(* IEC 61131-3 sources: JingjiangArm/moonboxpro_arm_8.4/Application/Application/任务列表/TensionTask/电机运动/MotionCtl_GantryTrap (part 2) *)

		//如果版辊周长变了/料膜厚度变了2023.12.27.171307
		IF (pstStGrpParam_Save^.rFilmThick_Confirm<>pstStGrpParam_Save^.rFilmThickNess_Using AND
			pstStGrpParam_Save^.rFilmThick_Confirm<>0 AND pstStGrpParam_Save^.rFilmThickNess_Using<>0) OR
			pstStUnitParam_Save^.rGirth_Confirmed_press_dn_NetRoller<>pstStUnitParam_Save^.rGirth_NetRoller OR
			pstStUnitParam_Save^.rGirth_Confirmed_press_dn_PrnRoller<>pstStUnitParam_Save^.rGirth_PrnRoller OR
			rGirth_PrnRoller_Mem <> pstStGrpParam_Save^.rGirth_PrnRoller THEN
			//处理一下位置更新2023.12.27.171801
			lrTemp:= g_rPos_press_dn_NetRoller_Pressure_MM*GC_LRMOTORPPR_TRAP*
						UINT_TO_REAL(pstStUnitParam_Save^.uiNum_NetRoller_Pressure)/
						pstStUnitParam_Save^.rScrewPitch_NetRoller_Pressure/
						UINT_TO_REAL(pstStUnitParam_Save^.uiDen_NetRoller_Pressure);

			IF i_pastStTrapAxisParam_Gantray^[2,iN].xRev_Motor_M THEN

				i_pastStTrapAxisParam_Gantray^[2,iN].lrposConfirm_Dn_Press_M:= i_pastStTrapAxisParam_Gantray^[2,iN].lrposConfirm_Dn_Press_M_Confirm-
						((
						(pstStGrpParam_Save^.rFilmThick_Manu-pstStGrpParam_Save^.rFilmThick_Confirm))*
						UINT_TO_LREAL(pstStUnitParam_Save^.uiNum_NetRoller_Pressure)*GC_LRMOTORPPR_TRAP/
						UINT_TO_LREAL(pstStUnitParam_Save^.uiDen_NetRoller_Pressure)/pstStUnitParam_Save^.rScrewPitch_NetRoller_Pressure);

				i_pastStTrapAxisParam_Gantray^[2,iN].lrposConfirm_Up_Press_M:= i_pastStTrapAxisParam_Gantray^[2,iN].lrposConfirm_Dn_Press_M-lrTemp;
			ELSE

					i_pastStTrapAxisParam_Gantray^[2,iN].lrposConfirm_Dn_Press_M:= i_pastStTrapAxisParam_Gantray^[2,iN].lrposConfirm_Dn_Press_M_Confirm+
						((
						(pstStGrpParam_Save^.rFilmThick_Manu-pstStGrpParam_Save^.rFilmThick_Confirm))*
						UINT_TO_LREAL(pstStUnitParam_Save^.uiNum_NetRoller_Pressure)*GC_LRMOTORPPR_TRAP/
						UINT_TO_LREAL(pstStUnitParam_Save^.uiDen_NetRoller_Pressure)/pstStUnitParam_Save^.rScrewPitch_NetRoller_Pressure);

				i_pastStTrapAxisParam_Gantray^[2,iN].lrposConfirm_Up_Press_M:= i_pastStTrapAxisParam_Gantray^[2,iN].lrposConfirm_Dn_Press_M+lrTemp;
			END_IF
			IF i_pastStTrapAxisParam_Gantray^[2,iN].xRev_Motor_G THEN

				i_pastStTrapAxisParam_Gantray^[2,iN].lrposConfirm_Dn_Press_G:= i_pastStTrapAxisParam_Gantray^[2,iN].lrposConfirm_Dn_Press_G_Confirm-
						(((*(i_pastStTrapAxisParam_Gantray^[2,iN].rweigth_Zero-
						i_pastStTrapAxisParam_Gantray^[2,iN].rweigth_Zero_Confirm)+*)
						(pstStGrpParam_Save^.rFilmThickNess_Using-pstStGrpParam_Save^.rFilmThick_Confirm))*
						UINT_TO_LREAL(pstStUnitParam_Save^.uiNum_NetRoller_Pressure)*GC_LRMOTORPPR_TRAP/
						UINT_TO_LREAL(pstStUnitParam_Save^.uiDen_NetRoller_Pressure)/pstStUnitParam_Save^.rScrewPitch_NetRoller_Pressure);
				i_pastStTrapAxisParam_Gantray^[2,iN].lrposConfirm_Up_Press_G:= i_pastStTrapAxisParam_Gantray^[2,iN].lrposConfirm_Dn_Press_G-lrTemp;
			ELSE

					i_pastStTrapAxisParam_Gantray^[2,iN].lrposConfirm_Dn_Press_G:= i_pastStTrapAxisParam_Gantray^[2,iN].lrposConfirm_Dn_Press_G_Confirm+
							(((i_pastStTrapAxisParam_Gantray^[2,iN].rweigth_Zero-
							i_pastStTrapAxisParam_Gantray^[2,iN].rweigth_Zero_Confirm)+
							(pstStGrpParam_Save^.rFilmThick_Manu-pstStGrpParam_Save^.rFilmThick_Confirm))*
							UINT_TO_LREAL(pstStUnitParam_Save^.uiNum_NetRoller_Pressure)*GC_LRMOTORPPR_TRAP/
							UINT_TO_LREAL(pstStUnitParam_Save^.uiDen_NetRoller_Pressure)/pstStUnitParam_Save^.rScrewPitch_NetRoller_Pressure);

				i_pastStTrapAxisParam_Gantray^[2,iN].lrposConfirm_Up_Press_G:= i_pastStTrapAxisParam_Gantray^[2,iN].lrposConfirm_Dn_Press_G+lrTemp;
			END_IF
			i_pastStTrapAxisParam_Gantray^[2,iN].lrposConfirm_Load_Unload_Press_M:= //换版位的物理位置是不变的2023.12.13.081145
				i_pastStTrapAxisParam_Gantray^[2,iN].lrposConfirm_Load_Unload_Press_M_Confirm;
			i_pastStTrapAxisParam_Gantray^[2,iN].lrposConfirm_Load_Unload_Press_G:=
				i_pastStTrapAxisParam_Gantray^[2,iN].lrposConfirm_Load_Unload_Press_G_Confirm;
		ELSE
			//bai.zy | 2024.03.21.130939 | 增加印刷位
			i_pastStTrapAxisParam_Gantray^[2,iN].lrposConfirm_Dn_Press_M:=
				i_pastStTrapAxisParam_Gantray^[2,iN].lrposConfirm_Dn_Press_M_Confirm;
			i_pastStTrapAxisParam_Gantray^[2,iN].lrposConfirm_Dn_Press_G:=
				i_pastStTrapAxisParam_Gantray^[2,iN].lrposConfirm_Dn_Press_G_Confirm;
			i_pastStTrapAxisParam_Gantray^[2,iN].lrposConfirm_Up_Press_M:=
				i_pastStTrapAxisParam_Gantray^[2,iN].lrposConfirm_Up_Press_M_Confirm;
			i_pastStTrapAxisParam_Gantray^[2,iN].lrposConfirm_Up_Press_G:=
				i_pastStTrapAxisParam_Gantray^[2,iN].lrposConfirm_Up_Press_G_Confirm;
			i_pastStTrapAxisParam_Gantray^[2,iN].lrposConfirm_Load_Unload_Press_M:= //换版位的物理位置是不变的2023.12.13.081145
				i_pastStTrapAxisParam_Gantray^[2,iN].lrposConfirm_Load_Unload_Press_M_Confirm;
			i_pastStTrapAxisParam_Gantray^[2,iN].lrposConfirm_Load_Unload_Press_G:=
				i_pastStTrapAxisParam_Gantray^[2,iN].lrposConfirm_Load_Unload_Press_G_Confirm;

		END_IF
	//2026.02.07.160105 计算网辊步进量

		afbKS_FB_GantryTrap_Calc_TargetPos_Net[iN](
			i_xEn:= TRUE,
			i_uiNum:= pstStUnitParam_Save^.uiNum_NetRoller_Pressure,
			i_uiDen:= pstStUnitParam_Save^.uiDen_NetRoller_Pressure,
			i_rScrewPitch:= pstStUnitParam_Save^.rScrewPitch_NetRoller_Pressure,
			i_rUp_Dn_Length:= g_rPos_press_dn_NetRoller_Pressure_MM,//1.35, //3mm
			i_rGirth_Roller:= pstStUnitParam_Save^.rGirth_NetRoller,
			i_xStopOrEstop_Valid:= xNeedMoveUp_Stop_Net,
			i_prGirth_Confirm:= ADR(pstStUnitParam_Save^.rGirth_Confirmed_press_dn_NetRoller),
			i_xFlag_Print:= pstStGrpParam_UnSave^.xFlag_Print,
			i_xStep_Fast:= pstStUnitParam_Save^.wFlag_PressFun.2,//^.xStep_Fast,
			i_rStep_Fast:= pstStGrpParam_Save^.rStep_Fast,
			i_rStep_Little:= pstStGrpParam_Save^.rStep_Little,
			i_rVel_Fast:= pstStGrpParam_Save^.rVel_Press_Net,//
			i_rVel_Little:= 0.1,
			i_plrTargetPos_All:= ADR(alrTargetPos_Net[iN]),
			i_plrTargetPos_M:= ADR(alrTargetPos_Net_M[iN]),
			i_plrTargetPos_G:= ADR(alrTargetPos_Net_G[iN]),
			i_pstStTrapAxisParam_Gantray:= ADR(i_pastStTrapAxisParam_Gantray^[2,iN]),
			i_xFlag_Estop:= i_xFlag_Estop,
			//i_rStep_HMI:= pstStUnitParam^.rStep_Pressure_Prn_Net,//2023.12.22.220303
			//i_rDistanceForAvoidPrnGear := 0,
			i_pxFinishConfirm_Adjust_PressDn := ADR(axFinishConfirm_Adjust_PressDn[iN]),//: POINTER TO BOOL;
			i_rStep_HMI_Use:=pstStUnitParam_Save^.rStep_Pressure_Prn_Net,
			i_rProportion:=1.0,
			i_xMove_to_Up_Estop := pstStGrpParam_Save^.wCtl_Pressure_Up_Dn.1,
			i_ReqResetEstop := i_ReqResetEstop,
			i_rMaxErr := rMaxErr,
			o_xEn=> ,
			o_rVel=> o_arVel_Net[iN],
			o_lrTargetPos_All=> o_alrTargetPos_Net[iN],
			o_lrTargetPos_M=> o_alrTargetPos_Net_M[iN],
			o_lrTargetPos_G=> o_alrTargetPos_Net_G[iN],
			o_lrTemp_Len_Up_Pos=>alrTemp_Len_Up_Pos_Net[iN],
			o_lrTemp_Len_Load_Unload_Pos=>alrTemp_Len_Load_Unload_Pos_Net[iN]);

		pstStUnitParam_Save^.rPos_load_unload_NetRoller_Pressure_M:=
			i_pastStTrapAxisParam_Gantray^[2,iN].lrposConfirm_Load_Unload_Press_M_Confirm;
		pstStUnitParam_Save^.rPos_load_unload_NetRoller_Pressure_G:=
			i_pastStTrapAxisParam_Gantray^[2,iN].lrposConfirm_Load_Unload_Press_G_Confirm;
		pstStUnitParam_Save^.rPos_press_up_NetRoller_Pressure_M:=
			i_pastStTrapAxisParam_Gantray^[2,iN].lrposConfirm_Up_Press_M_Confirm;
		pstStUnitParam_Save^.rPos_press_up_NetRoller_Pressure_G:=
			i_pastStTrapAxisParam_Gantray^[2,iN].lrposConfirm_Up_Press_G_Confirm;
		pstStUnitParam_Save^.rPos_press_dn_NetRoller_Pressure_M:=
			i_pastStTrapAxisParam_Gantray^[2,iN].lrposConfirm_Dn_Press_M_Confirm;
		pstStUnitParam_Save^.rPos_press_dn_NetRoller_Pressure_G:=
			i_pastStTrapAxisParam_Gantray^[2,iN].lrposConfirm_Dn_Press_G_Confirm;
		pstStUnitParam_UnSave^.rPos_NetRoller_Pressure_M:= LREAL_TO_REAL(i_pastStTrapAxisParam_Gantray^[2,iN].lrCurPos_mm_M);
		pstStUnitParam_UnSave^.rPos_NetRoller_Pressure_G:= LREAL_TO_REAL(i_pastStTrapAxisParam_Gantray^[2,iN].lrCurPos_mm_G);

		//bai.zy | 2024.01.15.105513 | 合压位换版位标定完成标志
		pstStUnitParam_Save^.xConfirmDnPosDne_NetRoller_Pressure_M := i_pastStTrapAxisParam_Gantray^[2,iN].xConfirmDnPosDne_Pressure_M;
		pstStUnitParam_Save^.xConfirmDnPosDne_NetRoller_Pressure_G := i_pastStTrapAxisParam_Gantray^[2,iN].xConfirmDnPosDne_Pressure_G;
		pstStUnitParam_Save^.xConfirmload_unloadPosDne_NetRoller_Pressure_M := i_pastStTrapAxisParam_Gantray^[2,iN].xConfirmload_unloadPosDne_Pressure_M;
		pstStUnitParam_Save^.xConfirmload_unloadPosDne_NetRoller_Pressure_G := i_pastStTrapAxisParam_Gantray^[2,iN].xConfirmload_unloadPosDne_Pressure_G;

		//2024.10.21.121704
		IF pstStUnitParam_UnSave^.xConfirmParallelPos_Net THEN//平行确认按钮
			pstStUnitParam_Save^.axPressLimit_Min[2] := TRUE;
			pstStUnitParam_Save^.lrEncPosParallel_Net_M:=i_pastStTrapAxisParam_Gantray^[2,iN].lrEncPosParallel_M;//平行编码器值
			pstStUnitParam_Save^.lrEncPosParallel_Net_G:=i_pastStTrapAxisParam_Gantray^[2,iN].lrEncPosParallel_G;
			pstStUnitParam_UnSave^.xConfirmParallelPos_Net := FALSE;
		END_IF
		pstStUnitParam_UnSave^.rParallelError_Net_MM := i_pastStTrapAxisParam_Gantray^[2,iN].lrParallelError_MM;
		pstStUnitParam_Save^.lrPrintPosOffsetDn_Net_M:=i_pastStTrapAxisParam_Gantray^[2,iN].lrPrintPosOffsetDn_M;//合压偏移量
		pstStUnitParam_Save^.lrPrintPosOffsetDn_Net_G:=i_pastStTrapAxisParam_Gantray^[2,iN].lrPrintPosOffsetDn_G;

		IF pstStUnitParam_UnSave^.axCalidPressLimit_Max[2] THEN
			pstStUnitParam_UnSave^.axCalidPressLimit_Max[2] := FALSE;
			pstStUnitParam_Save^.axPressLimit_Max[2] := TRUE;
			pstStUnitParam_Save^.lrEncPosLimit_Net_M_Max := i_pastStTrapAxisParam_Gantray^[2,iN].lrEncPosLimit_M_Max ;
			pstStUnitParam_Save^.lrEncPosLimit_Net_G_Max := i_pastStTrapAxisParam_Gantray^[2,iN].lrEncPosLimit_G_Max ;
		END_IF

	END_FOR

	//版周长

	rGirth_PrnRoller_Mem := pstStGrpParam_Save^.rGirth_PrnRoller;		//	秦华不需要了

	FOR iN:=1 TO i_iGrpUnitNum_Pu BY 1 DO
		IF axFlag_Mode_Calid[iN] THEN
			g_xModeCalibSwitch_Flag := TRUE;
			IF NOT i_xDebugMode THEN
				g_xModeCalibSwitch_Flag := FALSE;
			END_IF
			EXIT;
		ELSE
			g_xModeCalibSwitch_Flag := FALSE;
		END_IF
	END_FOR

	IF i_xDebugMode THEN
		FOR iN := 1 TO i_iGrpUnitNum_Pu BY 1 DO
			pstStUnitParam_Save:= ADR(i_pstStSysParam^.astStUnitParam_Save[iN]);
			pstStUnitParam_UnSave:= ADR(i_pstStSysParam^.astStUnitParam_UnSave[iN]);
			axTRIG_ResetFlag_FinishCalid[iN](CLK:=g_axResetFlag_FinishCalid[iN]);
			IF axTRIG_ResetFlag_FinishCalid[iN].Q THEN
				g_axResetFlag_FinishCalid[iN] := FALSE;

				pstStUnitParam_Save^.xConfirmDnPosDne_PrnRoller_Pressure_M:=FALSE;
				pstStUnitParam_Save^.xConfirmDnPosDne_PrnRoller_Pressure_G:=FALSE;
				pstStUnitParam_Save^.xConfirmDnPosDne_NetRoller_Pressure_M:=FALSE;
				pstStUnitParam_Save^.xConfirmDnPosDne_NetRoller_Pressure_G:=FALSE;
				pstStUnitParam_Save^.xConfirmload_unloadPosDne_PrnRoller_Pressure_M:=FALSE;
				pstStUnitParam_Save^.xConfirmload_unloadPosDne_PrnRoller_Pressure_G:=FALSE;
				pstStUnitParam_Save^.xConfirmload_unloadPosDne_NetRoller_Pressure_M:=FALSE;
				pstStUnitParam_Save^.xConfirmload_unloadPosDne_NetRoller_Pressure_G:=FALSE;

				pstStUnitParam_Save^.xConfirmDnPosDne_StrRoller_Pressure_M:=FALSE;
				pstStUnitParam_Save^.xConfirmDnPosDne_StrRoller_Pressure_G:=FALSE;
				//印版
				pstStUnitParam_Save^.rPos_load_unload_PrnRoller_Pressure_M := 0;//换版位
				pstStUnitParam_Save^.rPos_load_unload_PrnRoller_Pressure_G := 0;
				pstStUnitParam_Save^.rPos_press_up_PrnRoller_Pressure_M := 0;//离压位
				pstStUnitParam_Save^.rPos_press_up_PrnRoller_Pressure_G := 0;
				pstStUnitParam_Save^.rPos_press_dn_PrnRoller_Pressure_M := 0;//合压位
				pstStUnitParam_Save^.rPos_press_dn_PrnRoller_Pressure_G := 0;
				pstStUnitParam_Save^.liABSPos_Prn_M := 0;
				pstStUnitParam_Save^.liABSPos_Prn_G := 0;
				//网辊
				pstStUnitParam_Save^.rPos_load_unload_NetRoller_Pressure_M := 0;//换版位
				pstStUnitParam_Save^.rPos_load_unload_NetRoller_Pressure_G := 0;
				pstStUnitParam_Save^.rPos_press_up_NetRoller_Pressure_M := 0;//离压位
				pstStUnitParam_Save^.rPos_press_up_NetRoller_Pressure_G := 0;
				pstStUnitParam_Save^.rPos_press_dn_NetRoller_Pressure_M := 0;//合压位
				pstStUnitParam_Save^.rPos_press_dn_NetRoller_Pressure_G := 0;
				pstStUnitParam_Save^.liABSPos_Net_M := 0;
				pstStUnitParam_Save^.liABSPos_Net_G := 0;
				//张带
				pstStUnitParam_Save^.rPos_load_unload_StrRoller_Pressure_M := 0;//换版位
				pstStUnitParam_Save^.rPos_load_unload_StrRoller_Pressure_G := 0;
				pstStUnitParam_Save^.rPos_press_up_StrRoller_Pressure_M := 0;//离压位
				pstStUnitParam_Save^.rPos_press_up_StrRoller_Pressure_G := 0;
				pstStUnitParam_Save^.rPos_press_dn_StrRoller_Pressure_M := 0;//合压位
				pstStUnitParam_Save^.rPos_press_dn_StrRoller_Pressure_G := 0;
				pstStUnitParam_Save^.liABSPos_Str_M := 0;
				pstStUnitParam_Save^.liABSPos_Str_G := 0;

				FOR iM := 1 TO gc_iMax_PressureRoller_Unit BY 1 DO
					aitargetStation[2*iM-1] := (i_pastStTrapAxisParam_Gantray^[iM,iN].iStationId_M);
					aitargetStation[2*iM] := (i_pastStTrapAxisParam_Gantray^[iM,iN].iStationId_G);
					aliABSEncPos[2*iM-1] := 0;
					aliABSEncPos[2*iM] := 0;
				END_FOR
				//iRtn := GT_RN_SetTrapCoordinate(targetNum:= INT_TO_BYTE(gc_iMax_PressureRoller_Unit*2), targetStation:= ADR(abytargetStation), targetAxis:= ADR(aliABSEncPos));

				axAxisRev[1]:= i_pastStTrapAxisParam_Gantray^[1,iN].xRev_Motor_M;
				axAxisRev[2]:= i_pastStTrapAxisParam_Gantray^[1,iN].xRev_Motor_G;
				axAxisRev[3]:= i_pastStTrapAxisParam_Gantray^[2,iN].xRev_Motor_M;
				axAxisRev[4]:= i_pastStTrapAxisParam_Gantray^[2,iN].xRev_Motor_G;
				axAxisRev[5]:= i_pastStTrapAxisParam_Gantray^[3,iN].xRev_Motor_M;
				axAxisRev[6]:= i_pastStTrapAxisParam_Gantray^[3,iN].xRev_Motor_G;

				iRtn := KS_SetTrapCoordinate(
						i_xEn:= TRUE,
						i_iTarget_Num:= INT_TO_BYTE(gc_iMax_PressureRoller_Unit*2),
						i_paiTargetStationList:= ADR(aitargetStation),
						i_paliABSEncPos:= ADR(aliABSEncPos),
						i_paxAxisRev:= ADR(axAxisRev),
						i_pastStAxisIdListInf:= i_pastStAxisIdListInf,
						i_pastStGetMotionSts:= i_pastStGetMotionSts,
						i_pstStSysStationInf := i_pstStSysStationInf,
						i_pstStSysGantryAxisInf := i_pstStSysGantryAxisInf,
						ADR(g_alrCurrentAbsPos_Debug));

			END_IF
		END_FOR
	END_IF

(*
	FOR iN := 1 TO i_iGrpUnitNum_Pu BY 1 DO
		pstStUnitParam_Save:= ADR(i_pstStSysParam^.astStUnitParam_Save[iN]);
		pstStUnitParam_UnSave:= ADR(i_pstStSysParam^.astStUnitParam_UnSave[iN]);
		//印刷过程中矫正合压位是否要重新清零清规划？？？？
		//矫正后更新当前参数值
		//2025.08.28.152652 | 矫正增加对于压力电机的位置判断，之前做过判断，但是不再范围内的位置还是被矫正了，这里再次判断一下
		IF axFinishConfirm_Adjust_PressDn[iN] AND
			pstStUnitParam_Save^.xLinkage AND
			(i_pastStTrapAxisParam_Gantray^[1,iN].byCurPos_M = 1 OR
			i_pastStTrapAxisParam_Gantray^[1,iN].byCurPos_M = 2 OR
			i_pastStTrapAxisParam_Gantray^[1,iN].byCurPos_M = 3 ) AND
			(i_pastStTrapAxisParam_Gantray^[1,iN].byCurPos_G = 1 OR
			i_pastStTrapAxisParam_Gantray^[1,iN].byCurPos_G = 2 OR
			i_pastStTrapAxisParam_Gantray^[1,iN].byCurPos_G = 3 ) AND
			(i_pastStTrapAxisParam_Gantray^[2,iN].byCurPos_M = 1 OR
			i_pastStTrapAxisParam_Gantray^[2,iN].byCurPos_M = 2 OR
			i_pastStTrapAxisParam_Gantray^[2,iN].byCurPos_M = 3 ) AND
			(i_pastStTrapAxisParam_Gantray^[2,iN].byCurPos_G = 1 OR
			i_pastStTrapAxisParam_Gantray^[2,iN].byCurPos_G = 2 OR
			i_pastStTrapAxisParam_Gantray^[2,iN].byCurPos_G = 3 ) THEN

			axFinishConfirm_Adjust_PressDn[iN] := FALSE;

			alrTemp_Len_Up_Pos_Prn[iN] := g_rPos_press_dn_PrnRoller_Pressure_MM(*i_pstStSysParam^.rPos_press_dn_PrnRoller_Pressure_MM*)*
										pstStUnitParam_Save^.uiNum_PrnRoller_Pressure*GC_LRMOTORPPR_TRAP/
										pstStUnitParam_Save^.uiDen_PrnRoller_Pressure/pstStUnitParam_Save^.rScrewPitch_PrnRoller_Pressure;
			alrTemp_Len_Load_Unload_Pos_Prn[iN] :=g_rPos_press_dn_PrnRoller_Pressure_MM(*i_pstStSysParam^.rPos_load_unload_PrnRoller_Pressure_MM*)*
										pstStUnitParam_Save^.uiNum_PrnRoller_Pressure*GC_LRMOTORPPR_TRAP/
										pstStUnitParam_Save^.uiDen_PrnRoller_Pressure/pstStUnitParam_Save^.rScrewPitch_PrnRoller_Pressure;
			//印版
			iRtn := GTN_RN_GetAxisAbsPosEx(cardNum:= 1, axis:= 1, pPos:= ADR(g_liAbsPos_M), stationId:= i_pastStTrapAxisParam_Gantray^[1,iN].iStationId_M);
			iRtn := GTN_RN_GetAxisAbsPosEx(cardNum:= 1, axis:= 1, pPos:= ADR(g_liAbsPos_G), stationId:= i_pastStTrapAxisParam_Gantray^[1,iN].iStationId_G);
			pstStUnitParam_Save^.rPos_press_dn_PrnRoller_Pressure_M:= 1;//LINT_TO_LREAL(g_liAbsPos_M);
			pstStUnitParam_Save^.rPos_press_dn_PrnRoller_Pressure_G:= 1;//LINT_TO_LREAL(g_liAbsPos_G);
			pstStUnitParam_Save^.rPos_press_up_PrnRoller_Pressure_M:= pstStUnitParam_Save^.rPos_press_dn_PrnRoller_Pressure_M + alrTemp_Len_Up_Pos_Prn[iN];//1;//LINT_TO_LREAL(g_liAbsPos_M);
			pstStUnitParam_Save^.rPos_press_up_PrnRoller_Pressure_G:= pstStUnitParam_Save^.rPos_press_dn_PrnRoller_Pressure_G + alrTemp_Len_Up_Pos_Prn[iN];//1;//LINT_TO_LREAL(g_liAbsPos_G);
			pstStUnitParam_Save^.rPos_load_unload_PrnRoller_Pressure_M:= pstStUnitParam_Save^.rPos_press_dn_PrnRoller_Pressure_M + alrTemp_Len_Load_Unload_Pos_Prn[iN];//1;//LINT_TO_LREAL(g_liAbsPos_M);
			pstStUnitParam_Save^.rPos_load_unload_PrnRoller_Pressure_G:= pstStUnitParam_Save^.rPos_press_dn_PrnRoller_Pressure_G + alrTemp_Len_Load_Unload_Pos_Prn[iN];//1;//LINT_TO_LREAL(g_liAbsPos_G);
			iRtn := GT_RN_SetTrapCoordinate(targetNum:=1 , targetStation:=ADR(i_pastStTrapAxisParam_Gantray^[1,iN].iStationId_M),targetAxis:= ADR(g_liAbsPos_M));
			iRtn := GT_RN_SetTrapCoordinate(targetNum:=1 , targetStation:=ADR(i_pastStTrapAxisParam_Gantray^[1,iN].iStationId_G),targetAxis:= ADR(g_liAbsPos_G));
			pstStUnitParam_Save^.liABSPos_Prn_M := g_liAbsPos_M;
			pstStUnitParam_Save^.liABSPos_Prn_G := g_liAbsPos_G;
			//网辊
			iRtn := GTN_RN_GetAxisAbsPosEx(cardNum:= 1, axis:= 1, pPos:= ADR(g_liAbsPos_M), stationId:= i_pastStTrapAxisParam_Gantray^[2,iN].iStationId_M);
			iRtn := GTN_RN_GetAxisAbsPosEx(cardNum:= 1, axis:= 1, pPos:= ADR(g_liAbsPos_G), stationId:= i_pastStTrapAxisParam_Gantray^[2,iN].iStationId_G);
			pstStUnitParam_Save^.rPos_press_dn_NetRoller_Pressure_M:= 1;//LINT_TO_LREAL(g_liAbsPos_M);
			pstStUnitParam_Save^.rPos_press_dn_NetRoller_Pressure_G:= 1;//LINT_TO_LREAL(g_liAbsPos_G);
			pstStUnitParam_Save^.rPos_press_up_NetRoller_Pressure_M:= pstStUnitParam_Save^.rPos_press_dn_NetRoller_Pressure_M + alrTemp_Len_Up_Pos_Net[iN];//1;//LINT_TO_LREAL(g_liAbsPos_M);
			pstStUnitParam_Save^.rPos_press_up_NetRoller_Pressure_G:= pstStUnitParam_Save^.rPos_press_dn_NetRoller_Pressure_G + alrTemp_Len_Up_Pos_Net[iN];//1;//LINT_TO_LREAL(g_liAbsPos_G);
			pstStUnitParam_Save^.rPos_load_unload_NetRoller_Pressure_M:= pstStUnitParam_Save^.rPos_press_dn_NetRoller_Pressure_M + alrTemp_Len_Load_Unload_Pos_Net[iN];//1;//LINT_TO_LREAL(g_liAbsPos_M);
			pstStUnitParam_Save^.rPos_load_unload_NetRoller_Pressure_G:= pstStUnitParam_Save^.rPos_press_dn_NetRoller_Pressure_G + alrTemp_Len_Load_Unload_Pos_Net[iN];//1;//LINT_TO_LREAL(g_liAbsPos_G);
			iRtn := GT_RN_SetTrapCoordinate(targetNum:=1 , targetStation:=ADR(i_pastStTrapAxisParam_Gantray^[2,iN].iStationId_M),targetAxis:= ADR(g_liAbsPos_M));
			iRtn := GT_RN_SetTrapCoordinate(targetNum:=1 , targetStation:=ADR(i_pastStTrapAxisParam_Gantray^[2,iN].iStationId_G),targetAxis:= ADR(g_liAbsPos_G));
			pstStUnitParam_Save^.liABSPos_Net_M := g_liAbsPos_M;
			pstStUnitParam_Save^.liABSPos_Net_G := g_liAbsPos_G;

		END_IF
	END_FOR
*)
IF xtest4 THEN
	xtest4:=FALSE;
	iRtn := GTN_RN_ReadAbsEncPos(cardIndex:= 1, stationPhyId:=  113, encoder:= 1, pPos:= ADR(lrAbsPos1));
	iRtn := GTN_RN_ReadAbsEncPos(cardIndex:= 1, stationPhyId:=  129, encoder:= 1, pPos:= ADR(lrAbsPos2));
	iRtn := GTN_RN_ReadAbsEncPos(cardIndex:= 1, stationPhyId:=  145, encoder:= 1, pPos:= ADR(lrAbsPos3));
	iRtn := GTN_RN_ReadAbsEncPos(cardIndex:= 1, stationPhyId:=  161, encoder:= 1, pPos:= ADR(lrAbsPos4));
END_IF

// iRtn := GTN_RN_ReadAbsEncPos(cardIndex:= 1, stationPhyId:=  114, encoder:= 1, pPos:= ADR(lrAbsPos2));
// iRtn := GTN_RN_ReadAbsEncPos(cardIndex:= 1, stationPhyId:=  115, encoder:= 1, pPos:= ADR(lrAbsPos3));
 //iRtn := GTN_RN_ReadAbsEncPos(cardIndex:= 1, stationPhyId:=  116, encoder:= 1, pPos:= ADR(lrAbsPos4));
//
// iRtn := GTN_RN_ReadAbsEncPos(cardIndex:= 1, stationPhyId:=  129, encoder:= 1, pPos:= ADR(lrAbsPos5));
//  iRtn := GTN_RN_ReadAbsEncPos(cardIndex:= 1, stationPhyId:=  130, encoder:= 1, pPos:= ADR(lrAbsPos6));
//  iRtn := GTN_RN_ReadAbsEncPos(cardIndex:= 1, stationPhyId:=  131, encoder:= 1, pPos:= ADR(lrAbsPos7));
 // iRtn := GTN_RN_ReadAbsEncPos(cardIndex:= 1, stationPhyId:=  132, encoder:= 1, pPos:= ADR(lrAbsPos8));

END_IF

(* ---- KS_FB_AxisEnCtl_GantryTrap.st ---- *)
(*@CES
Name=KS_FB_AxisEnCtl_GantryTrap
Type=FunctionBlock
TypeGuid=6f9dac99-8de1-4efc-8465-68ac443b7d08
Guid=6adbed21-caa4-496e-a20b-968a8a51526d
HasDeclaration=True
HasImplementation=True
*)
{DECLARATION}
FUNCTION_BLOCK KS_FB_AxisEnCtl_GantryTrap
VAR_INPUT
	i_xEn: BOOL;
	i_iGrpId: INT;
	i_iGrpGantryTrapGroup_Num: INT;
	i_iGrpGantryTrapMotion_Num: INT;
	i_aiGrpGantryTrapMotion_StdList: ARRAY [1..MAX_STATION_NUM] OF INT;
	i_pstStSysParam: POINTER TO StSysParam;
	i_pastStAxisIdListInf :POINTER TO ARRAY [1..128] OF StAxisIdListInf;
	i_pastStMotorParam_GantryTrap: POINTER TO ARRAY [1..MAX_STATION_NUM] OF StMotorParam_GantryTrap;
END_VAR
VAR_OUTPUT
	o_iAxisId_Master: INT;
END_VAR
VAR
	iN: INT;
	iAxisId: INT;
	iTypeId: INT;
	iUnitId: INT;
	iCoreId: INT;
	iGroupId : INT;
	pstStGrpParam_Save: POINTER TO StGrpParam_Save;
	pstStGrpParam_UnSave: POINTER TO StGrpParam_UnSave;

END_VAR

{IMPLEMENTATION}
IF i_xEn THEN
	IF (i_iGrpId=1 OR i_iGrpId=2) AND
		i_iGrpGantryTrapGroup_Num >0 AND
		i_pstStSysParam<>0 AND
		i_pastStAxisIdListInf<>0 AND
		i_pastStMotorParam_GantryTrap<>0 THEN
		pstStGrpParam_Save:= ADR(i_pstStSysParam^.astStGrpParam_Save[i_iGrpId]);
		pstStGrpParam_UnSave:= ADR(i_pstStSysParam^.astStGrpParam_UnSave[i_iGrpId]);

		FOR iGroupId:=1 TO i_iGrpGantryTrapGroup_Num BY 1 DO
			CASE i_pastStMotorParam_GantryTrap^[iGroupId].iTypeId OF
			TYPE_UNIT_PRN_PRESS_MASTER:
				i_pastStMotorParam_GantryTrap^[iGroupId].xMoveEn := pstStGrpParam_Save^.wCtl_Pressure_Up_Dn.5;//g_axEn_Motor_Gantry[i_iGrpId];
							//i_pstStSysParam^.astStUnitParam_UnSave[i_pastStMotorParam_GantryTrap^[iGroupId].iUnitId].byEn_Motor_Pressure.0;
				i_pastStMotorParam_GantryTrap^[iGroupId].xMoveRev_M :=
									i_pstStSysParam^.astStUnitParam_UnSave[i_pastStMotorParam_GantryTrap^[iGroupId].iUnitId].xMotRev_PrnRoller_Pressure_M;
				i_pastStMotorParam_GantryTrap^[iGroupId].xMoveRev_G :=
									i_pstStSysParam^.astStUnitParam_UnSave[i_pastStMotorParam_GantryTrap^[iGroupId].iUnitId].xMotRev_PrnRoller_Pressure_G;

			TYPE_UNIT_NET_PRESS_MASTER:
				i_pastStMotorParam_GantryTrap^[iGroupId].xMoveEn := pstStGrpParam_Save^.wCtl_Pressure_Up_Dn.5;
							//i_pstStSysParam^.astStUnitParam_UnSave[i_pastStMotorParam_GantryTrap^[iGroupId].iUnitId].byEn_Motor_Pressure.1;
				i_pastStMotorParam_GantryTrap^[iGroupId].xMoveRev_M :=
									i_pstStSysParam^.astStUnitParam_UnSave[i_pastStMotorParam_GantryTrap^[iGroupId].iUnitId].xMotRev_NetRoller_Pressure_M;
				i_pastStMotorParam_GantryTrap^[iGroupId].xMoveRev_G :=
									i_pstStSysParam^.astStUnitParam_UnSave[i_pastStMotorParam_GantryTrap^[iGroupId].iUnitId].xMotRev_NetRoller_Pressure_G;
			TYPE_UNIT_STR_PRESS_MASTER:
				i_pastStMotorParam_GantryTrap^[iGroupId].xMoveEn := pstStGrpParam_Save^.wCtl_Pressure_Up_Dn.5;
							//i_pstStSysParam^.astStUnitParam_UnSave[i_pastStMotorParam_GantryTrap^[iGroupId].iUnitId].byEn_Motor_Pressure.2;
				i_pastStMotorParam_GantryTrap^[iGroupId].xMoveRev_M :=
									i_pstStSysParam^.astStUnitParam_UnSave[i_pastStMotorParam_GantryTrap^[iGroupId].iUnitId].xMotRev_StrRoller_Pressure_M;
				i_pastStMotorParam_GantryTrap^[iGroupId].xMoveRev_G :=
									i_pstStSysParam^.astStUnitParam_UnSave[i_pastStMotorParam_GantryTrap^[iGroupId].iUnitId].xMotRev_StrRoller_Pressure_G;

			END_CASE

(*
			KS_HY_GetAxisIdForMotByStation(
				i_aiGrpGantryTrapMotion_StdList[iN],
				ADR(iAxisId),
				ADR(iTypeId),
				ADR(iUnitId),
				ADR(iCoreId),
				i_pastStAxisIdListInf);
			CASE iTypeId OF
			TYPE_UNIT_PRN_PRESS_MASTER:
				i_pastStMotorParam_GantryTrap^[iN].xMoveEn := i_pstStSysParam^.astStUnitParam_UnSave[iUnitId].byEn_Motor_Pressure.0;
				i_pastStMotorParam_GantryTrap^[iN].xMoveRev := i_pstStSysParam^.astStUnitParam_UnSave[iUnitId].xMotRev_PrnRoller_Pressure_M;
			TYPE_UNIT_PRN_PRESS_M:
				i_pastStMotorParam_GantryTrap^[iN].xMoveEn := i_pstStSysParam^.astStUnitParam_UnSave[iUnitId].byEn_Motor_Pressure.0;
				i_pastStMotorParam_GantryTrap^[iN].xMoveRev := i_pstStSysParam^.astStUnitParam_UnSave[iUnitId].xMotRev_PrnRoller_Pressure_M;
			TYPE_UNIT_PRN_PRESS_G:
				i_pastStMotorParam_GantryTrap^[iN].xMoveEn := i_pstStSysParam^.astStUnitParam_UnSave[iUnitId].byEn_Motor_Pressure.1;
				i_pastStMotorParam_GantryTrap^[iN].xMoveRev := i_pstStSysParam^.astStUnitParam_UnSave[iUnitId].xMotRev_PrnRoller_Pressure_G;
			TYPE_UNIT_NET_PRESS_MASTER:
				i_pastStMotorParam_GantryTrap^[iN].xMoveEn := i_pstStSysParam^.astStUnitParam_UnSave[iUnitId].byEn_Motor_Pressure.2;
				i_pastStMotorParam_GantryTrap^[iN].xMoveRev := i_pstStSysParam^.astStUnitParam_UnSave[iUnitId].xMotRev_NetRoller_Pressure_M;
			TYPE_UNIT_NET_PRESS_M:
				i_pastStMotorParam_GantryTrap^[iN].xMoveEn := i_pstStSysParam^.astStUnitParam_UnSave[iUnitId].byEn_Motor_Pressure.2;
				i_pastStMotorParam_GantryTrap^[iN].xMoveRev := i_pstStSysParam^.astStUnitParam_UnSave[iUnitId].xMotRev_NetRoller_Pressure_M;
			TYPE_UNIT_NET_PRESS_G:
				i_pastStMotorParam_GantryTrap^[iN].xMoveEn := i_pstStSysParam^.astStUnitParam_UnSave[iUnitId].byEn_Motor_Pressure.3;
				i_pastStMotorParam_GantryTrap^[iN].xMoveRev := i_pstStSysParam^.astStUnitParam_UnSave[iUnitId].xMotRev_NetRoller_Pressure_G;
			TYPE_UNIT_STR_PRESS_MASTER:
				i_pastStMotorParam_GantryTrap^[iN].xMoveEn := i_pstStSysParam^.astStUnitParam_UnSave[iUnitId].byEn_Motor_Pressure.4;
				i_pastStMotorParam_GantryTrap^[iN].xMoveRev := i_pstStSysParam^.astStUnitParam_UnSave[iUnitId].xMotRev_StrRoller_Pressure_M;
			TYPE_UNIT_STR_PRESS_M:
				i_pastStMotorParam_GantryTrap^[iN].xMoveEn := i_pstStSysParam^.astStUnitParam_UnSave[iUnitId].byEn_Motor_Pressure.4;
				i_pastStMotorParam_GantryTrap^[iN].xMoveRev := i_pstStSysParam^.astStUnitParam_UnSave[iUnitId].xMotRev_StrRoller_Pressure_M;
			TYPE_UNIT_STR_PRESS_G:
				i_pastStMotorParam_GantryTrap^[iN].xMoveEn := i_pstStSysParam^.astStUnitParam_UnSave[iUnitId].byEn_Motor_Pressure.5;
				i_pastStMotorParam_GantryTrap^[iN].xMoveRev := i_pstStSysParam^.astStUnitParam_UnSave[iUnitId].xMotRev_StrRoller_Pressure_G;
			END_CASE
*)
		END_FOR
	END_IF
ELSE
	;
END_IF

(* ---- KS_FB_AxisPosCtl_GantryTrap.st ---- *)
(*@CES
Name=KS_FB_AxisPosCtl_GantryTrap
Type=FunctionBlock
TypeGuid=6f9dac99-8de1-4efc-8465-68ac443b7d08
Guid=58bb9038-ba9b-45e2-97ef-dcb3af1a4c94
HasDeclaration=True
HasImplementation=True
*)
{DECLARATION}
FUNCTION_BLOCK KS_FB_AxisPosCtl_GantryTrap
VAR_INPUT
	i_xEn: BOOL;
	i_iGrpId: INT;
	i_iGrpUnitNum_Pu : INT;
	i_iGrpGantryTrapGroup_Num: INT;
	i_iGrpGantryTrapMotion_Num: INT;
	i_aiGrpGantryTrapMotion_StdList: ARRAY [1..MAX_STATION_NUM] OF INT;
	i_pstStSysParam: POINTER TO StSysParam;
	i_pastStAxisIdListInf :POINTER TO ARRAY [1..128] OF StAxisIdListInf;
	i_pastStMotorParam_GantryTrap: POINTER TO ARRAY [1..MAX_STATION_NUM] OF StMotorParam_GantryTrap;

	i_arvel_UnitPressure_Prn:  ARRAY [1..MAX_UNIT_NUM] OF REAL;
	i_arvel_UnitPressure_Net:  ARRAY [1..MAX_UNIT_NUM] OF REAL;
	i_alrTargetPos_Prn:   ARRAY [1..MAX_UNIT_NUM] OF LREAL;
	i_alrTargetPos_Prn_M:   ARRAY [1..MAX_UNIT_NUM] OF LREAL;
	i_alrTargetPos_Prn_G:   ARRAY [1..MAX_UNIT_NUM] OF LREAL;
	i_alrTargetPos_Net:   ARRAY [1..MAX_UNIT_NUM] OF LREAL;
	i_alrTargetPos_Net_M:   ARRAY [1..MAX_UNIT_NUM] OF LREAL;
	i_alrTargetPos_Net_G:   ARRAY [1..MAX_UNIT_NUM] OF LREAL;
END_VAR
VAR_OUTPUT
END_VAR
VAR
	iN: INT;
	iAxisId: INT;
	iTypeId: INT;
	iUnitId: INT;
	iCoreId: INT;
	iGroupId : INT;
	pstStGrpParam_Save: POINTER TO StGrpParam_Save;
	pstStGrpParam_UnSave: POINTER TO StGrpParam_UnSave;

END_VAR

{IMPLEMENTATION}
IF i_xEn THEN
	IF (i_iGrpId=1 OR i_iGrpId=2) AND
		i_iGrpGantryTrapGroup_Num > 0 AND
		i_pstStSysParam<>0 AND
		i_pastStAxisIdListInf<>0 AND
		i_pastStMotorParam_GantryTrap<>0 THEN
		pstStGrpParam_Save:= ADR(i_pstStSysParam^.astStGrpParam_Save[i_iGrpId]);
		pstStGrpParam_UnSave:= ADR(i_pstStSysParam^.astStGrpParam_UnSave[i_iGrpId]);

		FOR iGroupId := 1 TO i_iGrpUnitNum_Pu BY 1 DO
			i_pastStMotorParam_GantryTrap^[iGroupId].diMax_Vel :=REAL_TO_DINT(i_arvel_UnitPressure_Prn[iGroupId]);
			i_pastStMotorParam_GantryTrap^[iGroupId].liTarget_Pos_All := LREAL_TO_LINT(i_alrTargetPos_Prn[iGroupId]);
			i_pastStMotorParam_GantryTrap^[iGroupId].diMain_Axis_Shift := LREAL_TO_DINT(i_alrTargetPos_Prn_M[iGroupId]);
			i_pastStMotorParam_GantryTrap^[iGroupId].diSecond_Axis_Shift := LREAL_TO_DINT(i_alrTargetPos_Prn_G[iGroupId]);

			i_pastStMotorParam_GantryTrap^[iGroupId+i_iGrpUnitNum_Pu].diMax_Vel :=REAL_TO_DINT(i_arvel_UnitPressure_Net[iGroupId]);
			i_pastStMotorParam_GantryTrap^[iGroupId+i_iGrpUnitNum_Pu].liTarget_Pos_All := LREAL_TO_LINT(i_alrTargetPos_Net[iGroupId]);
			i_pastStMotorParam_GantryTrap^[iGroupId+i_iGrpUnitNum_Pu].diMain_Axis_Shift := LREAL_TO_DINT(i_alrTargetPos_Net_M[iGroupId]);
			i_pastStMotorParam_GantryTrap^[iGroupId+i_iGrpUnitNum_Pu].diSecond_Axis_Shift := LREAL_TO_DINT(i_alrTargetPos_Net_G[iGroupId]);
		END_FOR

// 		FOR iGroupId:=1 TO i_iGrpGantryTrapGroup_Num BY 1 DO
// 			i_pastStMotorParam_GantryTrap^[iGroupId].diMax_Vel :=100;
// 			i_pastStMotorParam_GantryTrap^[iGroupId].liTarget_Pos_All := 1000000;
// 			i_pastStMotorParam_GantryTrap^[iGroupId].diMain_Axis_Shift := 500000;
// 			i_pastStMotorParam_GantryTrap^[iGroupId].diSecond_Axis_Shift := 100000;
// 		END_FOR
	END_IF
ELSE
	;
END_IF

(* ---- KS_FB_CacuHypotenuse_V3.st ---- *)
(*@CES
Name=KS_FB_CacuHypotenuse_V3
Type=FunctionBlock
TypeGuid=6f9dac99-8de1-4efc-8465-68ac443b7d08
Guid=f624852b-9183-4541-83cd-e00bb1937fb0
HasDeclaration=True
HasImplementation=True
*)
{DECLARATION}
FUNCTION_BLOCK KS_FB_CacuHypotenuse_V3
VAR_INPUT
		i_xEn:BOOL;
		i_rPrRoller_Girth0:REAL;//确认合压位时的版辊周长
		i_rPrRoller_Girth:REAL;
		i_rBrRoller_Girth:REAL;
		i_rFilmThick_Confirm:REAL;//标定合压位时的料膜厚度
		i_rFilmThickNess_Using:REAL;//现在的料膜厚度
		i_rFix_Horizontal_Edge_X:REAL;
END_VAR
VAR_OUTPUT
		o_rCathetus_diff:REAL;
END_VAR
VAR
		rPrRadius0:REAL;//确认合压位时的版辊半径
		rPrRadius:REAL;//换版后的版辊半径
		rBrRadius:REAL;
		rHypotenuse_L0:REAL;//换版前的斜边
		rHypotenuse_L1:REAL;//换版后的斜边
		rCathetus0:REAL;//换版前直角边
		rCathetus1:REAL;//换版后直角边
		rCathetus_diff:REAL;
END_VAR

{IMPLEMENTATION}
IF i_xEn THEN
	IF i_rPrRoller_Girth0 > 0.0 THEN
		rPrRadius0 :=  i_rPrRoller_Girth0/ (2 * gc_lrPI);
	END_IF
	IF i_rPrRoller_Girth> 0.0 THEN
		rPrRadius := i_rPrRoller_Girth / (2 * gc_lrPI);
	END_IF

	IF i_rBrRoller_Girth > 0.0 THEN
		rBrRadius := i_rBrRoller_Girth / (2 * gc_lrPI);
	END_IF

	rHypotenuse_L0:=rPrRadius0+rBrRadius+i_rFilmThick_Confirm;
	rCathetus0:=SQRT(ABS((rHypotenuse_L0*rHypotenuse_L0) -(i_rFix_Horizontal_Edge_X*i_rFix_Horizontal_Edge_X)) );
	rHypotenuse_L1:=rPrRadius+rBrRadius+i_rFilmThickNess_Using;
	rCathetus1:=SQRT(ABS((rHypotenuse_L1*rHypotenuse_L1) -(i_rFix_Horizontal_Edge_X*i_rFix_Horizontal_Edge_X)) );
	rCathetus_diff:=rCathetus1-rCathetus0; //换版前和换版后合压位置的竖直位置差 mm
	o_rCathetus_diff:=rCathetus_diff;

END_IF

(* ---- KS_FB_CalcuDisplayT.st ---- *)
(*@CES
Name=KS_FB_CalcuDisplayT
Type=FunctionBlock
TypeGuid=6f9dac99-8de1-4efc-8465-68ac443b7d08
Guid=554f8a16-8195-4e33-a33d-03d9edef6993
HasDeclaration=True
HasImplementation=True
*)
{DECLARATION}
FUNCTION_BLOCK KS_FB_CalcuDisplayT
VAR_INPUT
	i_xEn:BOOL;
	i_rPrRoller_Girth:REAL;
	i_rNrRoller_Girth:REAL;
	i_rBrnRoller_Girth:REAL;
	//i_rPos_press_dn_PrnRoller_Pressure_MM:REAL;
	i_rFix_Horizontal_Edge_X:REAL;
	i_lrCurPos_mm:REAL;
END_VAR
VAR_OUTPUT
	o_rHypotenuse:REAL;
END_VAR
VAR
	rPrRadius:REAL;
	rNrRadius:REAL;
	rBrRadius:REAL;
	rHypotenuse_L0:REAL;
	rCathetus_Basic: REAL;
	rHypotenuse_L1:REAL;//斜边
	rHypotenuse:REAL;//斜边
	rCathetus:REAL;
END_VAR

{IMPLEMENTATION}
IF i_xEn THEN
	IF i_rPrRoller_Girth > 0.0 THEN
		rPrRadius := i_rPrRoller_Girth / (2 * gc_lrPI);
	END_IF
	IF i_rNrRoller_Girth > 0.0 THEN
		rNrRadius := i_rNrRoller_Girth / (2 * gc_lrPI);
	END_IF

	IF i_rBrnRoller_Girth > 0.0 THEN
		rBrRadius := i_rBrnRoller_Girth / (2 * gc_lrPI);
	END_IF
	rHypotenuse_L0:=rPrRadius+rBrRadius; //计算原始斜边
	rCathetus_Basic:=SQRT(ABS((rHypotenuse_L0*rHypotenuse_L0) -(i_rFix_Horizontal_Edge_X*i_rFix_Horizontal_Edge_X)) );//原始竖直边
	rCathetus:=rCathetus_Basic+i_lrCurPos_mm;
	rHypotenuse_L1:=SQRT(ABS(rCathetus*rCathetus+i_rFix_Horizontal_Edge_X*i_rFix_Horizontal_Edge_X));
	rHypotenuse:=rHypotenuse_L1-rPrRadius-rBrRadius;
	o_rHypotenuse:=rHypotenuse;
END_IF

(* ---- KS_FB_CalcuHypotenuse.st ---- *)
(*@CES
Name=KS_FB_CalcuHypotenuse
Type=FunctionBlock
TypeGuid=6f9dac99-8de1-4efc-8465-68ac443b7d08
Guid=d24b6977-ace1-4b02-9c22-6ad4a97686d8
HasDeclaration=True
HasImplementation=True
*)
{DECLARATION}
FUNCTION_BLOCK KS_FB_CalcuHypotenuse
VAR_INPUT
	i_xEn:BOOL;
	i_rPrRoller_Girth:REAL;
	i_rNrRoller_Girth:REAL;
	i_rBrRoller_Girth:REAL;
	i_rPos_press_dn_PrnRoller_Pressure_MM:REAL;
	i_rFix_Horizontal_Edge_X:REAL;
END_VAR
VAR_OUTPUT
	o_rPos_press_dn_PrnRoller_Pressure_MM:REAL;
END_VAR
VAR
rPrRadius:REAL;
rNrRadius:REAL;
rBrRadius:REAL;
rHypotenuse_L0:REAL;
rHypotenuse:REAL;//斜边
rCathetus:REAL;//直角边
rPos_press_dn_PrnRoller_Pressure_MM:REAL;
END_VAR

{IMPLEMENTATION}
IF i_xEn THEN
	IF i_rPrRoller_Girth > 0.0 THEN
		rPrRadius := i_rPrRoller_Girth / (2 * gc_lrPI);
	END_IF
	IF i_rNrRoller_Girth > 0.0 THEN
		rNrRadius := i_rNrRoller_Girth / (2 * gc_lrPI);
	END_IF

	IF i_rBrRoller_Girth > 0.0 THEN
		rBrRadius := i_rBrRoller_Girth / (2 * gc_lrPI);
	END_IF
	rHypotenuse_L0:=rPrRadius+rBrRadius; //计算原始斜边
	rHypotenuse:=(*3*)g_rPos_press_dn_PrnRoller_Pressure_MM+rHypotenuse_L0;	//斜边
	rCathetus:=SQRT(ABS((rHypotenuse_L0*rHypotenuse_L0) -(i_rFix_Horizontal_Edge_X*i_rFix_Horizontal_Edge_X)) );//竖直边
	rPos_press_dn_PrnRoller_Pressure_MM:=ABS(SQRT(ABS(rHypotenuse*rHypotenuse-i_rFix_Horizontal_Edge_X*i_rFix_Horizontal_Edge_X))-rCathetus);
	o_rPos_press_dn_PrnRoller_Pressure_MM:=rPos_press_dn_PrnRoller_Pressure_MM;
ELSE
	o_rPos_press_dn_PrnRoller_Pressure_MM := i_rPos_press_dn_PrnRoller_Pressure_MM;
END_IF

(* ---- KS_FB_CalcuHypotenuse_V2.st ---- *)
(*@CES
Name=KS_FB_CalcuHypotenuse_V2
Type=FunctionBlock
TypeGuid=6f9dac99-8de1-4efc-8465-68ac443b7d08
Guid=a8a80304-7605-4c77-80a2-5631ceae8e52
HasDeclaration=True
HasImplementation=True
*)
{DECLARATION}
FUNCTION_BLOCK KS_FB_CalcuHypotenuse_V2
VAR_INPUT
	i_xEn:BOOL;
	i_rPrRoller_Girth:REAL;
	i_rNrRoller_Girth:REAL;
	i_rBrRoller_Girth:REAL;
	i_rPos_press_dn_PrnRoller_Pressure_MM:REAL;
	i_rFix_Horizontal_Edge_X:REAL;
	i_lrCurPos_mm : LREAL;
END_VAR
VAR_OUTPUT
	o_rProportion:REAL;
END_VAR
VAR
rPrRadius:REAL;
rNrRadius:REAL;
rBrRadius:REAL;
rHypotenuse_L0:REAL;
rHypotenuse:REAL;//斜边
rCathetus:REAL;//直角边
rPos_press_dn_PrnRoller_Pressure_MM:REAL;
END_VAR

{IMPLEMENTATION}
IF i_xEn THEN
	IF i_rPrRoller_Girth > 0.0 THEN
		rPrRadius := i_rPrRoller_Girth / (2 * gc_lrPI);
	END_IF
	IF i_rNrRoller_Girth > 0.0 THEN
		rNrRadius := i_rNrRoller_Girth / (2 * gc_lrPI);
	END_IF

	IF i_rBrRoller_Girth > 0.0 THEN
		rBrRadius := i_rBrRoller_Girth / (2 * gc_lrPI);
	END_IF
	rHypotenuse_L0:=rPrRadius+rBrRadius + i_lrCurPos_mm; //计算原始斜边
	rHypotenuse:=(*3*)i_rPos_press_dn_PrnRoller_Pressure_MM+rHypotenuse_L0;	//斜边
	rCathetus:=SQRT(ABS((rHypotenuse_L0*rHypotenuse_L0) -(i_rFix_Horizontal_Edge_X*i_rFix_Horizontal_Edge_X)) );//竖直边
	rPos_press_dn_PrnRoller_Pressure_MM:=ABS(SQRT(ABS(rHypotenuse*rHypotenuse-i_rFix_Horizontal_Edge_X*i_rFix_Horizontal_Edge_X))-rCathetus);
	o_rProportion := rPos_press_dn_PrnRoller_Pressure_MM/i_rPos_press_dn_PrnRoller_Pressure_MM;
ELSE
	o_rProportion := 1;
END_IF

(* ---- KS_FB_CheckServeOnDone_GantryTrap.st ---- *)
(*@CES
Name=KS_FB_CheckServeOnDone_GantryTrap
Type=FunctionBlock
TypeGuid=6f9dac99-8de1-4efc-8465-68ac443b7d08
Guid=d3768567-e4db-4539-97ab-c25a5fceb7f7
HasDeclaration=True
HasImplementation=True
*)
{DECLARATION}
FUNCTION_BLOCK KS_FB_CheckServeOnDone_GantryTrap
VAR_INPUT
	i_xEn: BOOL;
	i_iGrpGantryTrapGroup_Num : INT;
	i_iGrpGantryTrapMotion_Num: INT;
	i_aiGrpGantryTrapMotion_StdList: ARRAY [1..MAX_STATION_NUM] OF INT;
	i_pstStSysParam: POINTER TO StSysParam;
	i_pastStAxisIdListInf :POINTER TO ARRAY [1..128] OF StAxisIdListInf;
	i_pastStGetMotionSts: POINTER TO ARRAY [1..MAX_STATION_NUM] OF StGetMotionSts;
	i_pastStMotorParam_GantryTrap: POINTER TO ARRAY [1..MAX_STATION_NUM] OF StMotorParam_GantryTrap;
	i_xFlag_StopOrEStop : BOOL;
END_VAR
VAR_OUTPUT
	o_xEn : BOOL;
	o_xDone : BOOL;
	o_iErrNo : INT;
	o_iErrAxisId : INT;
	o_iErrTypeId : INT;
	o_iErrUnitId : INT;
	o_iErrCoreId : INT;
	o_iErrGroupId : INT;
END_VAR
VAR
	iN : INT;
	aiErrServoOn_Cnt : ARRAY [1..128] OF INT;
	iServoOnNum : INT;
	iNotNeedServoOnNum : INT;
END_VAR

{IMPLEMENTATION}
o_xEn := i_xEn;
o_iErrNo := 0;
o_iErrAxisId := 0;
o_iErrTypeId := 0;
o_iErrUnitId := 0;
o_iErrCoreId := 0;
iServoOnNum := 0;
iNotNeedServoOnNum := 0;
IF i_xEn THEN
	IF i_pstStSysParam <> 0 AND
		i_pastStAxisIdListInf <> 0 AND
		i_pastStGetMotionSts <> 0 AND
		i_pastStMotorParam_GantryTrap <> 0 THEN
		FOR iN := 1 TO i_iGrpGantryTrapGroup_Num BY 1 DO
			IF i_pastStMotorParam_GantryTrap^[iN].xMoveEn THEN
				IF (*i_pastStGetMotionSts^[(i_pastStMotorParam_GantryTrap^[iN].iCoreId -1) * gc_ResCount_Profile + i_pastStMotorParam_GantryTrap^[iN].iAxisId].dwDriverSts.1 AND *)
					i_pastStGetMotionSts^[(i_pastStMotorParam_GantryTrap^[iN].iCoreId -1) * gc_ResCount_Profile + i_pastStMotorParam_GantryTrap^[iN].iAxisId].dwMotionSts.9 THEN
					iServoOnNum := iServoOnNum + 1;

					aiErrServoOn_Cnt[iN] := 0;
				ELSE
					aiErrServoOn_Cnt[iN] := aiErrServoOn_Cnt[iN] + 1;
					IF aiErrServoOn_Cnt[iN] > 10*1000/gc_TENSION_TSK_CYCLE_TIME THEN
						aiErrServoOn_Cnt[iN] := aiErrServoOn_Cnt[iN] -1;
// 						KS_HY_GetAxisIdForMotByStation(
// 							i_aiGrpGantryTrapMotion_StdList[iN],
// 							ADR(o_iErrAxisId),
// 							ADR(o_iErrTypeId),
// 							ADR(o_iErrUnitId),
// 							ADR(o_iErrCoreId),
// 							ADR(o_iErrGroupId),
// 							i_pastStAxisIdListInf);
						o_iErrAxisId := i_pastStMotorParam_GantryTrap^[iN].iAxisId;
						o_iErrTypeId := i_pastStMotorParam_GantryTrap^[iN].iTypeId;
						o_iErrUnitId := i_pastStMotorParam_GantryTrap^[iN].iUnitId;
						o_iErrCoreId := i_pastStMotorParam_GantryTrap^[iN].iCoreId;
						o_iErrGroupId := i_pastStMotorParam_GantryTrap^[iN].iGroupId;;
						o_iErrNo := -1;
					END_IF
					o_xDone := FALSE;
					EXIT;
				END_IF
			ELSE
				iNotNeedServoOnNum := iNotNeedServoOnNum + 1;
			END_IF
		END_FOR

		IF iServoOnNum = (i_iGrpGantryTrapGroup_Num - iNotNeedServoOnNum) THEN
			o_xDone := TRUE;
		END_IF
	END_IF
ELSE
	;
END_IF

(* ---- KS_FB_GantryTrap_Calc_TargetPos.st ---- *)
(*@CES
Name=KS_FB_GantryTrap_Calc_TargetPos
Type=FunctionBlock
TypeGuid=6f9dac99-8de1-4efc-8465-68ac443b7d08
Guid=0bce8d11-2bc3-4a0c-8964-1d70c50dfb2a
HasDeclaration=True
HasImplementation=True
*)
{DECLARATION}
FUNCTION_BLOCK KS_FB_GantryTrap_Calc_TargetPos
//一组龙门的控制？
VAR_INPUT
	i_xEn: BOOL;
	i_uiNum: UINT;//压力电机减速比
	i_uiDen: UINT;
	i_rScrewPitch: REAL;//压力电机螺杆螺距
	i_rUp_Dn_Length: REAL;//合压位离压位距离
	i_rGirth_Roller: REAL;//棍子周长，秦华记录带长，只对于张带辊有效
	i_xStopOrEstop_Valid: BOOL;

	i_prGirth_Confirm: POINTER TO REAL;//记录标定的周长
	i_xFlag_Print: BOOL;
	i_xStep_Fast: BOOL;//长步选择
	i_rStep_Fast: REAL;//长步步幅
	i_rStep_Little: REAL;//长步步幅
	i_rVel_Fast: REAL;//快速
	i_rVel_Little: REAL;//慢速
	i_plrTargetPos_All: POINTER TO LREAL;
	i_plrTargetPos_M: POINTER TO LREAL;
	i_plrTargetPos_G: POINTER TO LREAL;

	i_pstStTrapAxisParam_Gantray : POINTER TO StTrapAxisParam_Gantray;
	i_xFlag_Estop: BOOL;
//	i_rDistanceForAvoidPrnGear: REAL;
	i_pxFinishConfirm_Adjust_PressDn : POINTER TO BOOL;
	//2026.01.16.140531  新增品字型
	i_rStep_HMI_Use: REAL;
	i_rProportion :REAL;
	i_xMove_to_Up_Estop : BOOL;
	i_ReqResetEstop: BOOL;//急停复位
	i_rMaxErr : REAL;

END_VAR
VAR_OUTPUT
	o_xEn: BOOL;
	o_rVel: REAL;
	o_lrTargetPos_All: LREAL;
	o_lrTargetPos_M: LREAL;
	o_lrTargetPos_G: LREAL;
	o_lrTemp_Len_Up_Pos : LREAL;
	o_lrTemp_Len_Load_Unload_Pos : LREAL;
	//2026.01.17.93413 新增
	o_lrK_Dynamic:LREAL;
END_VAR
VAR
	//根据版周长和标定位置计算出对应版周的对应位置
// 	lrposConfirm_Dn_Press_Temp_M:LREAL;//合压位标定；
// 	lrposConfirm_Up_Press_Temp_M:LREAL;//离压位标定；
// 	lrposConfirm_Load_Unload_Press_Temp_M:LREAL;//换版位标定；
// 	lrposConfirm_Dn_Press_Temp_G:LREAL;//合压位标定；
// 	lrposConfirm_Up_Press_Temp_G:LREAL;//离压位标定；
// 	lrposConfirm_Load_Unload_Press_Temp_G:LREAL;//换版位标定；
	lrTemp: LREAL;
	fbTRIG_Confirm_load_unload: R_TRIG;
	fbTRIG_Confirm_PressUp: R_TRIG;
	fbTRIG_Confirm_PressDn: R_TRIG;
	fbTRIG_Confirm_ParallelPos: R_TRIG;
	fbTRIG_xCalidPressLimit_Max: R_TRIG;
	lrTemp_Len_Load_Unload_Pos: LREAL;
	lrTemp_100um_pos:LREAL:=167772;
	xPosIn: BOOL;
	xPosOut: BOOL;
	rStep_Use: REAL;
	xClearVelSetCurPos_For: BOOL;
	iClearVelSetCurPosCount_For:INT;
	xClearVelSetCurPos_Rev: BOOL;
	iClearVelSetCurPosCount_Rev:INT;
	rTemp_MovePos_M: REAL;
	rTemp_MovePos_G: REAL;
	lrTarPos_M_Temp: LREAL;
	lrTarPos_G_Temp: LREAL;
	xClearVelSetCurPos_HandWheel: BOOL;
	iClearVelSetCurPosCount_HandWheel:INT;
	rTemp: REAL;
	xPreStop_Prf_M: BOOL;
	xPreStop_Prf_G: BOOL;
	xMove_TO_TarFlag_M: BOOL;
	xMove_TO_TarFlag_G: BOOL;

	lrEncParallelError_M : LREAL;
	lrEncParallelError_G : LREAL;

	rStep_Panel : REAL;
	rVel_Panel : REAL;

	lrK_Dynamic:REAL:=1;
//	lrDistanceForAvoidPrnGear : LREAL;
	fbTRIG_Move_to_Up: R_TRIG;
	fbTRIG_Move_to_Dn: R_TRIG;
	fbTRIG_Move_to_Unload: R_TRIG;

	//2026.05.10.003923 | + | 增加限位保护
	rLast_TarPos_All : REAL;
	rLast_TarPos_M : REAL;
	rLast_TarPos_G : REAL;
	rLast_ErrPos : REAL;

	rErr_TarPos_All : REAL;
	rErr_TarPos_M : REAL;
	rErr_TarPos_G : REAL;
	rErr_Pos : REAL;

END_VAR

{IMPLEMENTATION}
IF i_xEn THEN
	IF i_uiNum<>0 AND i_uiDen<>0 AND i_rScrewPitch<>0 AND i_pstStTrapAxisParam_Gantray<>0 THEN
//2023.12.27.185420处理都放外面
		//先计算当前位置（M侧和G侧）//先就以合压位作为原点吧

// 			g_rtest:=i_rVel_Fast;
// 			g_uitest1:=i_uiNum;
// 			g_uitest2:=i_uiDen;
// 			g_rtest1:=i_rScrewPitch;

		i_pstStTrapAxisParam_Gantray^.lrPos_ZeroPos_Enc_M:= i_pstStTrapAxisParam_Gantray^.lrposConfirm_Dn_Press_M;
		IF i_pstStTrapAxisParam_Gantray^.lrPos_ZeroPos_Enc_M<>0 THEN//未标定
			//当前位置需要根据电机正反计算
			IF i_pstStTrapAxisParam_Gantray^.xRev_Motor_M THEN
				i_pstStTrapAxisParam_Gantray^.lrCurPos_mm_M:= -1*
					(i_pstStTrapAxisParam_Gantray^.lrPos_CurPos_Enc_M-i_pstStTrapAxisParam_Gantray^.lrPos_ZeroPos_Enc_M)*
					i_rScrewPitch*UINT_TO_LREAL(i_uiDen)/GC_LRMOTORPPR_TRAP/UINT_TO_REAL(i_uiNum);
				//计算一下前后表面的位置

			ELSE
				i_pstStTrapAxisParam_Gantray^.lrCurPos_mm_M:= 1*
					(i_pstStTrapAxisParam_Gantray^.lrPos_CurPos_Enc_M-i_pstStTrapAxisParam_Gantray^.lrPos_ZeroPos_Enc_M)*
					i_rScrewPitch*UINT_TO_LREAL(i_uiDen)/GC_LRMOTORPPR_TRAP/UINT_TO_REAL(i_uiNum);
			END_IF
		ELSE
			i_pstStTrapAxisParam_Gantray^.lrCurPos_mm_M:= 0;
		END_IF
		//i_pstStTrapAxisParam_Gantray^.lrPos_ZeroPos_Enc_G:= i_pstStTrapAxisParam_Gantray^.lrposConfirm_Dn_Press_G_Confirm;
		i_pstStTrapAxisParam_Gantray^.lrPos_ZeroPos_Enc_G:= i_pstStTrapAxisParam_Gantray^.lrposConfirm_Dn_Press_G;
		IF i_pstStTrapAxisParam_Gantray^.lrPos_ZeroPos_Enc_G<>0 THEN//未标定
			//当前位置需要根据电机正反计算
			IF i_pstStTrapAxisParam_Gantray^.xRev_Motor_G THEN
				i_pstStTrapAxisParam_Gantray^.lrCurPos_mm_G:= -1*
					(i_pstStTrapAxisParam_Gantray^.lrPos_CurPos_Enc_G-i_pstStTrapAxisParam_Gantray^.lrPos_ZeroPos_Enc_G)*
					i_rScrewPitch*UINT_TO_LREAL(i_uiDen)/GC_LRMOTORPPR_TRAP/UINT_TO_REAL(i_uiNum);
			ELSE
				i_pstStTrapAxisParam_Gantray^.lrCurPos_mm_G:= 1*
					(i_pstStTrapAxisParam_Gantray^.lrPos_CurPos_Enc_G-i_pstStTrapAxisParam_Gantray^.lrPos_ZeroPos_Enc_G)*
					i_rScrewPitch*UINT_TO_LREAL(i_uiDen)/GC_LRMOTORPPR_TRAP/UINT_TO_REAL(i_uiNum);
			END_IF
		ELSE
			i_pstStTrapAxisParam_Gantray^.lrCurPos_mm_G:= 0;
		END_IF

		//处理一下当前位置判断
		i_pstStTrapAxisParam_Gantray^.byCurPos_M:= 0;
		lrTemp_100um_pos:= 0.1*GC_LRMOTORPPR_TRAP*
						UINT_TO_REAL(i_uiNum)/
						i_rScrewPitch/
						UINT_TO_REAL(i_uiDen);
		IF i_pstStTrapAxisParam_Gantray^.xRev_Motor_M THEN
			IF (i_pstStTrapAxisParam_Gantray^.lrPos_CurPos_Enc_M - i_pstStTrapAxisParam_Gantray^.lrposConfirm_Dn_Press_M)>lrTemp_100um_pos THEN
				(*版辊操作侧位置在合压位和底辊中间*)
				i_pstStTrapAxisParam_Gantray^.byCurPos_M:= 1;
			ELSIF (i_pstStTrapAxisParam_Gantray^.lrPos_CurPos_Enc_M - i_pstStTrapAxisParam_Gantray^.lrposConfirm_Dn_Press_M)>(-1*lrTemp_100um_pos) AND
				(i_pstStTrapAxisParam_Gantray^.lrPos_CurPos_Enc_M - i_pstStTrapAxisParam_Gantray^.lrposConfirm_Dn_Press_M)<lrTemp_100um_pos THEN
				(*在合压位*)
				i_pstStTrapAxisParam_Gantray^.byCurPos_M:= 2;
			ELSIF  (i_pstStTrapAxisParam_Gantray^.lrPos_CurPos_Enc_M - i_pstStTrapAxisParam_Gantray^.lrposConfirm_Dn_Press_M)<(-1*lrTemp_100um_pos) AND
				(i_pstStTrapAxisParam_Gantray^.lrPos_CurPos_Enc_M - i_pstStTrapAxisParam_Gantray^.lrposConfirm_Up_Press_M)>lrTemp_100um_pos THEN
				(*在合压位和离压位之间*)
				i_pstStTrapAxisParam_Gantray^.byCurPos_M:= 3;
			ELSIF (i_pstStTrapAxisParam_Gantray^.lrPos_CurPos_Enc_M - i_pstStTrapAxisParam_Gantray^.lrposConfirm_Up_Press_M)>(-1*lrTemp_100um_pos) AND
				(i_pstStTrapAxisParam_Gantray^.lrPos_CurPos_Enc_M - i_pstStTrapAxisParam_Gantray^.lrposConfirm_Up_Press_M)<lrTemp_100um_pos THEN
				(*在离压位*)
				i_pstStTrapAxisParam_Gantray^.byCurPos_M:= 4;
			ELSIF  (i_pstStTrapAxisParam_Gantray^.lrPos_CurPos_Enc_M - i_pstStTrapAxisParam_Gantray^.lrposConfirm_Up_Press_M)<(-1*lrTemp_100um_pos) AND
				(i_pstStTrapAxisParam_Gantray^.lrPos_CurPos_Enc_M - i_pstStTrapAxisParam_Gantray^.lrposConfirm_Load_Unload_Press_M)>lrTemp_100um_pos THEN
				(*在换版位和离压位之间*)
				i_pstStTrapAxisParam_Gantray^.byCurPos_M:= 5;
			ELSE(*其他都算在换版位*)
				i_pstStTrapAxisParam_Gantray^.byCurPos_M:= 0;
			END_IF
		ELSE
			IF (i_pstStTrapAxisParam_Gantray^.lrPos_CurPos_Enc_M - i_pstStTrapAxisParam_Gantray^.lrposConfirm_Dn_Press_M)<(-1*lrTemp_100um_pos) THEN
				(*版辊操作侧位置在合压位和底辊中间*)
				i_pstStTrapAxisParam_Gantray^.byCurPos_M:= 1;
			ELSIF (i_pstStTrapAxisParam_Gantray^.lrPos_CurPos_Enc_M - i_pstStTrapAxisParam_Gantray^.lrposConfirm_Dn_Press_M)>(-1*lrTemp_100um_pos) AND
				(i_pstStTrapAxisParam_Gantray^.lrPos_CurPos_Enc_M - i_pstStTrapAxisParam_Gantray^.lrposConfirm_Dn_Press_M)<lrTemp_100um_pos THEN
				(*在合压位*)
				i_pstStTrapAxisParam_Gantray^.byCurPos_M:= 2;
			ELSIF  (i_pstStTrapAxisParam_Gantray^.lrPos_CurPos_Enc_M - i_pstStTrapAxisParam_Gantray^.lrposConfirm_Up_Press_M)<(-1*lrTemp_100um_pos) AND
				(i_pstStTrapAxisParam_Gantray^.lrPos_CurPos_Enc_M - i_pstStTrapAxisParam_Gantray^.lrposConfirm_Dn_Press_M)>lrTemp_100um_pos THEN
				(*在合压位和离压位之间*)
				i_pstStTrapAxisParam_Gantray^.byCurPos_M:= 3;
			ELSIF (i_pstStTrapAxisParam_Gantray^.lrPos_CurPos_Enc_M - i_pstStTrapAxisParam_Gantray^.lrposConfirm_Up_Press_M)>(-1*lrTemp_100um_pos) AND
				(i_pstStTrapAxisParam_Gantray^.lrPos_CurPos_Enc_M - i_pstStTrapAxisParam_Gantray^.lrposConfirm_Up_Press_M)<lrTemp_100um_pos THEN
				(*在离压位*)
				i_pstStTrapAxisParam_Gantray^.byCurPos_M:= 4;
			ELSIF  (i_pstStTrapAxisParam_Gantray^.lrPos_CurPos_Enc_M - i_pstStTrapAxisParam_Gantray^.lrposConfirm_Load_Unload_Press_M)<(-1*lrTemp_100um_pos) AND
				(i_pstStTrapAxisParam_Gantray^.lrPos_CurPos_Enc_M - i_pstStTrapAxisParam_Gantray^.lrposConfirm_Up_Press_M)>lrTemp_100um_pos THEN
				(*在换版位和离压位之间*)
				i_pstStTrapAxisParam_Gantray^.byCurPos_M:= 5;
			ELSE(*其他都算在换版位*)
				i_pstStTrapAxisParam_Gantray^.byCurPos_M:= 0;
			END_IF
		END_IF
		i_pstStTrapAxisParam_Gantray^.byCurPos_G:= 0;
		lrTemp_100um_pos:= 0.1*GC_LRMOTORPPR_TRAP*
						UINT_TO_REAL(i_uiNum)/
						i_rScrewPitch/
						UINT_TO_REAL(i_uiDen);
		IF i_pstStTrapAxisParam_Gantray^.xRev_Motor_G THEN
			IF (i_pstStTrapAxisParam_Gantray^.lrPos_CurPos_Enc_G - i_pstStTrapAxisParam_Gantray^.lrposConfirm_Dn_Press_G)>lrTemp_100um_pos THEN
				(*版辊操作侧位置在合压位和底辊中间*)
				i_pstStTrapAxisParam_Gantray^.byCurPos_G:= 1;
			ELSIF (i_pstStTrapAxisParam_Gantray^.lrPos_CurPos_Enc_G - i_pstStTrapAxisParam_Gantray^.lrposConfirm_Dn_Press_G)>(-1*lrTemp_100um_pos) AND
				(i_pstStTrapAxisParam_Gantray^.lrPos_CurPos_Enc_G - i_pstStTrapAxisParam_Gantray^.lrposConfirm_Dn_Press_G)<lrTemp_100um_pos THEN
				(*在合压位*)
				i_pstStTrapAxisParam_Gantray^.byCurPos_G:= 2;
			ELSIF  (i_pstStTrapAxisParam_Gantray^.lrPos_CurPos_Enc_G - i_pstStTrapAxisParam_Gantray^.lrposConfirm_Dn_Press_G)<(-1*lrTemp_100um_pos) AND
				(i_pstStTrapAxisParam_Gantray^.lrPos_CurPos_Enc_G - i_pstStTrapAxisParam_Gantray^.lrposConfirm_Up_Press_G)>lrTemp_100um_pos THEN
				(*在合压位和离压位之间*)
				i_pstStTrapAxisParam_Gantray^.byCurPos_G:= 3;
			ELSIF (i_pstStTrapAxisParam_Gantray^.lrPos_CurPos_Enc_G - i_pstStTrapAxisParam_Gantray^.lrposConfirm_Up_Press_G)>(-1*lrTemp_100um_pos) AND
				(i_pstStTrapAxisParam_Gantray^.lrPos_CurPos_Enc_G - i_pstStTrapAxisParam_Gantray^.lrposConfirm_Up_Press_G)<lrTemp_100um_pos THEN
				(*在离压位*)
				i_pstStTrapAxisParam_Gantray^.byCurPos_G:= 4;
			ELSIF  (i_pstStTrapAxisParam_Gantray^.lrPos_CurPos_Enc_G - i_pstStTrapAxisParam_Gantray^.lrposConfirm_Up_Press_G)<(-1*lrTemp_100um_pos) AND
				(i_pstStTrapAxisParam_Gantray^.lrPos_CurPos_Enc_G - i_pstStTrapAxisParam_Gantray^.lrposConfirm_Load_Unload_Press_G)>lrTemp_100um_pos THEN
				(*在换版位和离压位之间*)
				i_pstStTrapAxisParam_Gantray^.byCurPos_G:= 5;
			ELSE(*其他都算在换版位*)
				i_pstStTrapAxisParam_Gantray^.byCurPos_G:= 0;
			END_IF
		ELSE
			IF (i_pstStTrapAxisParam_Gantray^.lrPos_CurPos_Enc_G - i_pstStTrapAxisParam_Gantray^.lrposConfirm_Dn_Press_G)<(-1*lrTemp_100um_pos) THEN
				(*版辊操作侧位置在合压位和底辊中间*)
				i_pstStTrapAxisParam_Gantray^.byCurPos_G:= 1;
			ELSIF (i_pstStTrapAxisParam_Gantray^.lrPos_CurPos_Enc_G - i_pstStTrapAxisParam_Gantray^.lrposConfirm_Dn_Press_G)>(-1*lrTemp_100um_pos) AND
				(i_pstStTrapAxisParam_Gantray^.lrPos_CurPos_Enc_G - i_pstStTrapAxisParam_Gantray^.lrposConfirm_Dn_Press_G)<lrTemp_100um_pos THEN
				(*在合压位*)
				i_pstStTrapAxisParam_Gantray^.byCurPos_G:= 2;
			ELSIF  (i_pstStTrapAxisParam_Gantray^.lrPos_CurPos_Enc_G - i_pstStTrapAxisParam_Gantray^.lrposConfirm_Up_Press_G)<(-1*lrTemp_100um_pos) AND
				(i_pstStTrapAxisParam_Gantray^.lrPos_CurPos_Enc_G - i_pstStTrapAxisParam_Gantray^.lrposConfirm_Dn_Press_G)>lrTemp_100um_pos THEN
				(*在合压位和离压位之间*)
				i_pstStTrapAxisParam_Gantray^.byCurPos_G:= 3;
			ELSIF (i_pstStTrapAxisParam_Gantray^.lrPos_CurPos_Enc_G - i_pstStTrapAxisParam_Gantray^.lrposConfirm_Up_Press_G)>(-1*lrTemp_100um_pos) AND
				(i_pstStTrapAxisParam_Gantray^.lrPos_CurPos_Enc_G - i_pstStTrapAxisParam_Gantray^.lrposConfirm_Up_Press_G)<lrTemp_100um_pos THEN
				(*在离压位*)
				i_pstStTrapAxisParam_Gantray^.byCurPos_G:= 4;
			ELSIF  (i_pstStTrapAxisParam_Gantray^.lrPos_CurPos_Enc_G - i_pstStTrapAxisParam_Gantray^.lrposConfirm_Load_Unload_Press_G)<(-1*lrTemp_100um_pos) AND
				(i_pstStTrapAxisParam_Gantray^.lrPos_CurPos_Enc_G - i_pstStTrapAxisParam_Gantray^.lrposConfirm_Up_Press_G)>lrTemp_100um_pos THEN
				(*在换版位和离压位之间*)
				i_pstStTrapAxisParam_Gantray^.byCurPos_G:= 5;
			ELSE(*其他都算在换版位*)
				i_pstStTrapAxisParam_Gantray^.byCurPos_G:= 0;
			END_IF

		END_IF

		//这里处理一下再次按按钮逻辑-运行过程中不能再动了
		IF i_pstStTrapAxisParam_Gantray^.xMove_To_Dn_Press_ing AND
			i_pstStTrapAxisParam_Gantray^.byCurPos_G=2 AND
			i_pstStTrapAxisParam_Gantray^.byCurPos_M=2 THEN//到位了，就可以处理其他按钮
			i_pstStTrapAxisParam_Gantray^.xMove_To_Dn_Press_ing:= FALSE;
			i_pstStTrapAxisParam_Gantray^.xMove_To_Dn_Press_end:= TRUE;

		END_IF
		IF i_pstStTrapAxisParam_Gantray^.xMove_To_Up_Press_ing AND
			i_pstStTrapAxisParam_Gantray^.byCurPos_G=4 AND
			i_pstStTrapAxisParam_Gantray^.byCurPos_M=4 THEN//到位了，就可以处理其他按钮
			i_pstStTrapAxisParam_Gantray^.xMove_To_Up_Press_ing:= FALSE;
		END_IF
		IF i_pstStTrapAxisParam_Gantray^.xMove_To_Load_Unload_Press_ing AND
			i_pstStTrapAxisParam_Gantray^.byCurPos_G=0 AND
			i_pstStTrapAxisParam_Gantray^.byCurPos_M=0 THEN//到位了，就可以处理其他按钮
			i_pstStTrapAxisParam_Gantray^.xMove_To_Load_Unload_Press_ing:= FALSE;
		END_IF

		fbTRIG_Move_to_Up(CLK:= i_pstStTrapAxisParam_Gantray^.xMove_To_Up_Press_ing);
		fbTRIG_Move_to_Dn(CLK:= i_pstStTrapAxisParam_Gantray^.xMove_To_Dn_Press_ing);
		fbTRIG_Move_to_Unload(CLK:= i_pstStTrapAxisParam_Gantray^.xMove_To_Load_Unload_Press_ing);
		IF fbTRIG_Move_to_Up.Q OR fbTRIG_Move_to_Dn.Q OR fbTRIG_Move_to_Unload.Q THEN
			xMove_TO_TarFlag_M:= FALSE;
			xMove_TO_TarFlag_G:= FALSE;
		END_IF

		IF xPreStop_Prf_M<>i_pstStTrapAxisParam_Gantray^.xAxisPrfStop_M THEN
			IF i_pstStTrapAxisParam_Gantray^.xAxisPrfStop_M THEN
				xMove_TO_TarFlag_M:= TRUE;
			ELSE
				xMove_TO_TarFlag_M:= FALSE;
			END_IF
			xPreStop_Prf_M:= i_pstStTrapAxisParam_Gantray^.xAxisPrfStop_M;
		END_IF
		IF xPreStop_Prf_G<>i_pstStTrapAxisParam_Gantray^.xAxisPrfStop_G THEN
			IF i_pstStTrapAxisParam_Gantray^.xAxisPrfStop_G THEN
				xMove_TO_TarFlag_G:= TRUE;
			ELSE
				xMove_TO_TarFlag_G:= FALSE;
			END_IF
			xPreStop_Prf_G:= i_pstStTrapAxisParam_Gantray^.xAxisPrfStop_G;
		END_IF

		IF (i_pstStTrapAxisParam_Gantray^.xMove_To_Load_Unload_Press_ing OR
			i_pstStTrapAxisParam_Gantray^.xMove_To_Up_Press_ing OR
			i_pstStTrapAxisParam_Gantray^.xMove_To_Dn_Press_ing) THEN
			i_pstStTrapAxisParam_Gantray^.xMove_To_PressUp:= FALSE;
			i_pstStTrapAxisParam_Gantray^.xMove_To_Load_Unload:= FALSE;
			i_pstStTrapAxisParam_Gantray^.xMove_To_PressDn:= FALSE;
			i_xStopOrEstop_Valid:= FALSE;
		END_IF

		IF (xMove_TO_TarFlag_M AND xMove_TO_TarFlag_G) AND
			(i_pstStTrapAxisParam_Gantray^.xMove_To_Load_Unload_Press_ing OR
			i_pstStTrapAxisParam_Gantray^.xMove_To_Up_Press_ing OR
			i_pstStTrapAxisParam_Gantray^.xMove_To_Dn_Press_ing) THEN
			i_pstStTrapAxisParam_Gantray^.xMove_To_Load_Unload_Press_ing:= FALSE;
			i_pstStTrapAxisParam_Gantray^.xMove_To_Up_Press_ing:= FALSE;
			i_pstStTrapAxisParam_Gantray^.xMove_To_Dn_Press_ing:= FALSE;
// 			xMove_TO_TarFlag_G:= FALSE;
// 			xMove_TO_TarFlag_M:= FALSE;
		END_IF
//bai.zy | 2024.01.15.101452 | 标定完成标志
		IF i_pstStTrapAxisParam_Gantray^.xConfirmDnPosDne_Pressure_M AND i_pstStTrapAxisParam_Gantray^.xConfirmDnPosDne_Pressure_G THEN

			xPosIn:= FALSE;
			xPosOut:= FALSE;
			IF i_pstStTrapAxisParam_Gantray^.byCurPos_M=0 AND i_pstStTrapAxisParam_Gantray^.byCurPos_G=0 THEN
				IF i_pstStTrapAxisParam_Gantray^.xMove_To_PressUp THEN
					xPosIn:= TRUE;
					xPosOut:= FALSE;
				END_IF
			ELSIF i_pstStTrapAxisParam_Gantray^.byCurPos_M=4 AND i_pstStTrapAxisParam_Gantray^.byCurPos_G=4 THEN
				IF i_pstStTrapAxisParam_Gantray^.xMove_To_Load_Unload THEN
					xPosIn:= FALSE;
					xPosOut:= TRUE;
				END_IF
				IF i_pstStTrapAxisParam_Gantray^.xMove_To_PressDn THEN
					xPosIn:= TRUE;
					xPosOut:= FALSE;
					i_pstStTrapAxisParam_Gantray^.xCanReFlashPos := TRUE;
					i_pstStTrapAxisParam_Gantray^.xRefleshPos := FALSE;
				END_IF
			ELSIF i_pstStTrapAxisParam_Gantray^.byCurPos_M=5 AND i_pstStTrapAxisParam_Gantray^.byCurPos_G=5 THEN
				IF i_pstStTrapAxisParam_Gantray^.xMove_To_PressUp THEN
					xPosIn:= TRUE;
					xPosOut:= FALSE;
				END_IF
				IF i_pstStTrapAxisParam_Gantray^.xMove_To_Load_Unload THEN
					xPosIn:= FALSE;
					xPosOut:= TRUE;
				END_IF
			ELSIF (i_pstStTrapAxisParam_Gantray^.byCurPos_M=1 OR
					i_pstStTrapAxisParam_Gantray^.byCurPos_M=2 OR
					i_pstStTrapAxisParam_Gantray^.byCurPos_M=3) AND
				 (i_pstStTrapAxisParam_Gantray^.byCurPos_G=1 OR
					i_pstStTrapAxisParam_Gantray^.byCurPos_G=2 OR
					i_pstStTrapAxisParam_Gantray^.byCurPos_G=3) THEN
				IF i_pstStTrapAxisParam_Gantray^.xMove_To_PressUp OR i_xStopOrEstop_Valid OR i_ReqResetEstop THEN//liya
					xPosIn:= FALSE;
					xPosOut:= TRUE;
					i_pstStTrapAxisParam_Gantray^.xRefleshPos := TRUE;
				END_IF
				IF i_pstStTrapAxisParam_Gantray^.xMove_To_PressDn THEN//heya
					xPosIn:= TRUE;
					xPosOut:= FALSE;
				END_IF
			END_IF
		ELSE
			xPosIn:= FALSE;
			xPosOut:= FALSE;
			i_pstStTrapAxisParam_Gantray^.xCanReFlashPos := FALSE;
			i_pstStTrapAxisParam_Gantray^.xRefleshPos := FALSE;
			i_pstStTrapAxisParam_Gantray^.xMove_To_PressDn := FALSE;
			i_pstStTrapAxisParam_Gantray^.xMove_To_PressUp := FALSE;
			i_pstStTrapAxisParam_Gantray^.xMove_To_Load_Unload := FALSE;
		END_IF
		//处理界面按钮

		//IF i_xStep_Fast THEN
//2026.04.09.225246这里不能再算步进量了，会有误动作的2026.04.09.225309
(*			rStep_Use:= i_rVel_Fast*GC_LRMOTORPPR_TRAP*
					UINT_TO_REAL(i_uiNum)/
					i_rScrewPitch/
					UINT_TO_REAL(i_uiDen);//为了方便这里直接换算成脉冲吧
*)			o_rVel:= i_rVel_Fast*GC_LRMOTORPPR_TRAP*
					UINT_TO_REAL(i_uiNum)/
					i_rScrewPitch/
					UINT_TO_REAL(i_uiDen)/1000.0;

// 		ELSE
// //				rStep_Use:= i_rStep_Little/5.0*2.0*GC_LRMOTORPPR_TRAP;
// //				o_arVel[iN]:= i_rVel_Little/5.0 *2.0*GC_LRMOTORPPR_TRAP/1000.0;
// 			rStep_Use:= i_rStep_Little*GC_LRMOTORPPR_TRAP*
// 					UINT_TO_REAL(i_uiNum)/
// 					i_rScrewPitch/
// 					UINT_TO_REAL(i_uiDen);//为了方便这里直接换算成脉冲吧
// 			o_rVel:= i_rVel_Little*GC_LRMOTORPPR_TRAP*
// 					UINT_TO_REAL(i_uiNum)/
// 					i_rScrewPitch/
// 					UINT_TO_REAL(i_uiDen)/1000.0;
//		END_IF
//bai.zy | 2024.01.05.104330 | 手轮与界面操作冲突
(*2026.04.09.235930
		IF NOT (i_pstStTrapAxisParam_Gantray^.xMoveRev_Long OR
			i_pstStTrapAxisParam_Gantray^.xMoveFor_Long OR
			i_pstStTrapAxisParam_Gantray^.xMove_To_Load_Unload_Press_ing OR
			i_pstStTrapAxisParam_Gantray^.xMove_To_Up_Press_ing OR
			i_pstStTrapAxisParam_Gantray^.xMove_To_Dn_Press_ing) THEN
*)
			rStep_Use:= i_rStep_HMI_Use*GC_LRMOTORPPR_TRAP*i_rProportion*
				UINT_TO_REAL(i_uiNum)/
				i_rScrewPitch/
				UINT_TO_REAL(i_uiDen);
			o_rVel:= i_rVel_Fast*GC_LRMOTORPPR_TRAP*
				UINT_TO_REAL(i_uiNum)/
				i_rScrewPitch/
				UINT_TO_REAL(i_uiDen)/1000.0;

			//2026.01.16.153921
(*
		ELSE
			;
		END_IF
*)
		IF i_pstStTrapAxisParam_Gantray^.xMoveFor_M	THEN
			i_plrTargetPos_M^:= i_plrTargetPos_M^+(-1*rStep_Use);
		ELSIF i_pstStTrapAxisParam_Gantray^.xMoveRev_M THEN
			i_plrTargetPos_M^:= i_plrTargetPos_M^+(1*rStep_Use);
		END_IF
		IF i_pstStTrapAxisParam_Gantray^.xMoveFor_G	THEN
			i_plrTargetPos_G^:= i_plrTargetPos_G^+(-1*rStep_Use);
		ELSIF i_pstStTrapAxisParam_Gantray^.xMoveRev_G THEN
			i_plrTargetPos_G^:= i_plrTargetPos_G^+(1*rStep_Use);
		END_IF

		rTemp:= (g_rTest_StepLength/1000.0)*GC_LRMOTORPPR_TRAP*
					UINT_TO_REAL(i_uiNum)/
					i_rScrewPitch/
					UINT_TO_REAL(i_uiDen);//为了方便这里直接换算成脉冲吧

		IF i_pstStTrapAxisParam_Gantray^.xMoveFor_Test_For_Rev_For THEN
			i_plrTargetPos_All^:= i_plrTargetPos_All^+(-1*rTemp);
		ELSIF i_pstStTrapAxisParam_Gantray^.xMoveFor_Test_For_Rev_Rev THEN
			i_plrTargetPos_All^:= i_plrTargetPos_All^+(1*rTemp);
		END_IF
//2024.12.03.152342 | 增加调试阶段测试压力电机反复来回运行
		IF i_pstStTrapAxisParam_Gantray^.xPressDebugMode_MoveFor THEN
			rTemp := ((i_pstStTrapAxisParam_Gantray^.lrEncPosParallel_M - i_pstStTrapAxisParam_Gantray^.lrPos_CurPos_Enc_M)+
						(i_pstStTrapAxisParam_Gantray^.lrEncPosParallel_G - i_pstStTrapAxisParam_Gantray^.lrPos_CurPos_Enc_G))/2;

			o_rVel:= i_rVel_Fast*GC_LRMOTORPPR_TRAP*
				UINT_TO_REAL(i_uiNum)/
				i_rScrewPitch/
				UINT_TO_REAL(i_uiDen)/1000.0;

			i_plrTargetPos_All^:= i_plrTargetPos_All^+(1*rTemp);
		ELSIF i_pstStTrapAxisParam_Gantray^.xPressDebugMode_MoveRev THEN
			rTemp := ((i_pstStTrapAxisParam_Gantray^.lrEncPosLimit_M_Max - i_pstStTrapAxisParam_Gantray^.lrPos_CurPos_Enc_M)+
						(i_pstStTrapAxisParam_Gantray^.lrEncPosLimit_G_Max - i_pstStTrapAxisParam_Gantray^.lrPos_CurPos_Enc_G))/2;
			o_rVel:= i_rVel_Fast*GC_LRMOTORPPR_TRAP*
				UINT_TO_REAL(i_uiNum)/
				i_rScrewPitch/
				UINT_TO_REAL(i_uiDen)/1000.0;

			i_plrTargetPos_All^:= i_plrTargetPos_All^+(1*rTemp);
		END_IF

		//2023.11.29.182021在这里处理一下避让吧
		IF i_pstStTrapAxisParam_Gantray^.xMove_To_Up_Avoidance AND
			(NOT i_pstStTrapAxisParam_Gantray^.xMove_To_Up_Avoidance_ing) AND
			 (i_pstStTrapAxisParam_Gantray^.byCurPos_M=1 OR
				i_pstStTrapAxisParam_Gantray^.byCurPos_M=2 OR
				i_pstStTrapAxisParam_Gantray^.byCurPos_M=3) AND
			 (i_pstStTrapAxisParam_Gantray^.byCurPos_G=1 OR
				i_pstStTrapAxisParam_Gantray^.byCurPos_G=2 OR
				i_pstStTrapAxisParam_Gantray^.byCurPos_G=3) THEN
			i_pstStTrapAxisParam_Gantray^.xMove_To_Up_Avoidance_ing:= TRUE;
			i_plrTargetPos_All^:= i_plrTargetPos_All^+i_pstStTrapAxisParam_Gantray^.rMoveUp_mm_Avoidance*GC_LRMOTORPPR_TRAP*
					UINT_TO_REAL(i_uiNum)/
					i_rScrewPitch/
					UINT_TO_REAL(i_uiDen);
		END_IF
		IF i_pstStTrapAxisParam_Gantray^.xMove_To_Up_Avoidance_ing AND
			i_pstStTrapAxisParam_Gantray^.xMove_To_Dn_Avoidance THEN
			i_pstStTrapAxisParam_Gantray^.xMove_To_Up_Avoidance_ing:= FALSE;
			i_plrTargetPos_All^:= i_plrTargetPos_All^-i_pstStTrapAxisParam_Gantray^.rMoveUp_mm_Avoidance*GC_LRMOTORPPR_TRAP*
					UINT_TO_REAL(i_uiNum)/
					i_rScrewPitch/
					UINT_TO_REAL(i_uiDen);
		END_IF
		IF i_pstStTrapAxisParam_Gantray^.xRollerMoveFor THEN
			i_plrTargetPos_All^:= i_plrTargetPos_All^+(-1*rStep_Use);
		ELSIF i_pstStTrapAxisParam_Gantray^.xRollerMoveRev THEN
			i_plrTargetPos_All^:= i_plrTargetPos_All^+(1*rStep_Use);
		END_IF
		IF i_pstStTrapAxisParam_Gantray^.xMoveFor_Long THEN
			i_plrTargetPos_All^:= i_plrTargetPos_All^+(-1*rStep_Use)*gc_TENSION_TSK_CYCLE_TIME*2/1000.0;
			iClearVelSetCurPosCount_For:= 0;
			//xClearVelSetCurPos_For:= FALSE;
			xClearVelSetCurPos_For:= TRUE;
		ELSE
			//xClearVelSetCurPos_For:= TRUE;
			IF xClearVelSetCurPos_For THEN
				o_rVel:= 0;
				iClearVelSetCurPosCount_For:= iClearVelSetCurPosCount_For+1;
				IF iClearVelSetCurPosCount_For>=3 THEN
					xClearVelSetCurPos_For:= FALSE;
					iClearVelSetCurPosCount_For:= 0;
					IF i_pstStTrapAxisParam_Gantray^.xRev_Motor_M THEN(*bai.zy | 2024.07.04.153851 | 加0.5丝补偿，电机停止效果更好*)
						i_plrTargetPos_All^:= -i_pstStTrapAxisParam_Gantray^.lrPos_CurPos_Prf+0.05*lrTemp_100um_pos;
					ELSE
						i_plrTargetPos_All^:= i_pstStTrapAxisParam_Gantray^.lrPos_CurPos_Prf-0.05*lrTemp_100um_pos;
					END_IF
// 				ELSE
// 					IF i_pstStTrapAxisParam_Gantray^.xRev_Motor_M THEN
// 						i_plrTargetPos_All^:= -i_pstStTrapAxisParam_Gantray^.lrPos_CurPos_Prf;
// 					ELSE
// 						i_plrTargetPos_All^:= i_pstStTrapAxisParam_Gantray^.lrPos_CurPos_Prf;
// 					END_IF
				END_IF
			END_IF
		END_IF
		IF i_pstStTrapAxisParam_Gantray^.xMoveRev_Long THEN
			i_plrTargetPos_All^:= i_plrTargetPos_All^+(1*rStep_Use)*gc_TENSION_TSK_CYCLE_TIME*2/1000.0;
			iClearVelSetCurPosCount_Rev:= 0;
			//xClearVelSetCurPos_Rev:= FALSE;
			xClearVelSetCurPos_Rev:= TRUE;
		ELSE
			//xClearVelSetCurPos_Rev:= TRUE;
			IF xClearVelSetCurPos_Rev THEN
				o_rVel:= 0;
				iClearVelSetCurPosCount_Rev:= iClearVelSetCurPosCount_Rev+1;
				IF iClearVelSetCurPosCount_Rev>=3 THEN
					xClearVelSetCurPos_Rev:= FALSE;
					iClearVelSetCurPosCount_Rev:= 0;
					IF i_pstStTrapAxisParam_Gantray^.xRev_Motor_M THEN(*bai.zy | 2024.07.04.153851 | 加0.5丝补偿，电机停止效果更好*)
						i_plrTargetPos_All^:= -i_pstStTrapAxisParam_Gantray^.lrPos_CurPos_Prf+0.05*lrTemp_100um_pos;
					ELSE														(**)
						i_plrTargetPos_All^:= i_pstStTrapAxisParam_Gantray^.lrPos_CurPos_Prf-0.05*lrTemp_100um_pos;
					END_IF
// 				ELSE
// 					IF i_pstStTrapAxisParam_Gantray^.xRev_Motor_M THEN
// 						i_plrTargetPos_All^:= -i_pstStTrapAxisParam_Gantray^.lrPos_CurPos_Prf;
// 					ELSE
// 						i_plrTargetPos_All^:= i_pstStTrapAxisParam_Gantray^.lrPos_CurPos_Prf;
// 					END_IF
				END_IF
			END_IF
		END_IF
		IF ( i_pstStTrapAxisParam_Gantray^.xMove_To_Load_Unload OR
			i_pstStTrapAxisParam_Gantray^.xMove_To_PressUp OR
			i_pstStTrapAxisParam_Gantray^.xMove_To_PressDn OR i_xStopOrEstop_Valid OR i_ReqResetEstop) THEN//前往换版位
			o_rVel:= i_rVel_Fast*GC_LRMOTORPPR_TRAP*
					UINT_TO_REAL(i_uiNum)/
					i_rScrewPitch/
					UINT_TO_REAL(i_uiDen)/1000.0;

// 			g_rtest:=i_rVel_Fast;
// 			g_uitest1:=i_uiNum;
// 			g_uitest2:=i_uiDen;
// 			g_rtest1:=i_rScrewPitch;
//2026.04.13.03357|在一个不规范的位置，操作了离合压或者换版，没有方向信号，清除标志，不进入运行状态置位
			IF (NOT xPosIn) AND (NOT xPosOut) THEN
				i_pstStTrapAxisParam_Gantray^.xMove_To_Load_Unload:= FALSE;
				i_pstStTrapAxisParam_Gantray^.xMove_To_PressUp:= FALSE;
				i_pstStTrapAxisParam_Gantray^.xMove_To_PressDn:= FALSE;
				i_xStopOrEstop_Valid:= FALSE;
			END_IF
//2026.04.13.03525
			IF i_pstStTrapAxisParam_Gantray^.xMove_To_Load_Unload  THEN
				i_pstStTrapAxisParam_Gantray^.xMove_To_Load_Unload_Press_ing:= TRUE;
				lrTarPos_M_Temp:= i_pstStTrapAxisParam_Gantray^.lrposConfirm_Load_Unload_Press_M;
				lrTarPos_G_Temp:= i_pstStTrapAxisParam_Gantray^.lrposConfirm_Load_Unload_Press_G;

			ELSIF (i_pstStTrapAxisParam_Gantray^.xMove_To_PressUp OR i_xStopOrEstop_Valid OR i_ReqResetEstop) AND(NOT i_pstStTrapAxisParam_Gantray^.xMove_To_Up_Press_ing) THEN
				IF (i_pstStTrapAxisParam_Gantray^.byCurPos_M=0 OR
					i_pstStTrapAxisParam_Gantray^.byCurPos_M=1 OR
					i_pstStTrapAxisParam_Gantray^.byCurPos_M=2 OR
					i_pstStTrapAxisParam_Gantray^.byCurPos_M=3) AND
					(i_pstStTrapAxisParam_Gantray^.byCurPos_G=0 OR
					i_pstStTrapAxisParam_Gantray^.byCurPos_G=1 OR
					i_pstStTrapAxisParam_Gantray^.byCurPos_G=2 OR
					i_pstStTrapAxisParam_Gantray^.byCurPos_G=3) THEN
						i_pstStTrapAxisParam_Gantray^.xMove_To_Up_Press_ing:= TRUE;
						i_pstStTrapAxisParam_Gantray^.xMove_To_Dn_Press_end:= FALSE;
							lrTarPos_M_Temp:= i_pstStTrapAxisParam_Gantray^.lrposConfirm_Up_Press_M;
							lrTarPos_G_Temp:= i_pstStTrapAxisParam_Gantray^.lrposConfirm_Up_Press_G;
				END_IF

			ELSIF i_pstStTrapAxisParam_Gantray^.xMove_To_PressDn AND (NOT i_pstStTrapAxisParam_Gantray^.xMove_To_Dn_Press_ing) THEN
				i_pstStTrapAxisParam_Gantray^.xMove_To_Dn_Press_ing:= TRUE;

				lrTarPos_M_Temp:= i_pstStTrapAxisParam_Gantray^.lrposConfirm_Dn_Press_M;
				lrTarPos_G_Temp:= i_pstStTrapAxisParam_Gantray^.lrposConfirm_Dn_Press_G;

			END_IF
			rTemp_MovePos_M:= ABS(lrTarPos_M_Temp-
				i_pstStTrapAxisParam_Gantray^.lrPos_CurPos_Enc_M);
			rTemp_MovePos_G:= ABS(lrTarPos_G_Temp-
				i_pstStTrapAxisParam_Gantray^.lrPos_CurPos_Enc_G);

		//2026.03.28.16390	test
// 			IF i_pstStTrapAxisParam_Gantray^.xMove_To_PressDn OR i_pstStTrapAxisParam_Gantray^.xMove_To_PressUp THEN
// 				g_lrtest1:=lrTarPos_M_Temp;
// 				g_lrtest2:=i_pstStTrapAxisParam_Gantray^.lrPos_CurPos_Enc_M;
// 				g_lrtest3:=lrTarPos_G_Temp;
// 				g_lrtest4:=i_pstStTrapAxisParam_Gantray^.lrPos_CurPos_Enc_G;
// 			END_IF

			IF xPosOut THEN
				IF rTemp_MovePos_M=rTemp_MovePos_G THEN
					i_plrTargetPos_All^:= i_plrTargetPos_All^+rTemp_MovePos_M;
				ELSIF rTemp_MovePos_M>rTemp_MovePos_G THEN
					i_plrTargetPos_All^:= i_plrTargetPos_All^+(rTemp_MovePos_G);
					i_plrTargetPos_M^:= i_plrTargetPos_M^+(rTemp_MovePos_M-rTemp_MovePos_G);
				ELSIF rTemp_MovePos_M<rTemp_MovePos_G THEN
					i_plrTargetPos_All^:= i_plrTargetPos_All^+(rTemp_MovePos_M);
					i_plrTargetPos_G^:= i_plrTargetPos_G^+(rTemp_MovePos_G-rTemp_MovePos_M);
				END_IF
			ELSIF xPosIn THEN
				IF rTemp_MovePos_M=rTemp_MovePos_G THEN
					i_plrTargetPos_All^:= i_plrTargetPos_All^-rTemp_MovePos_M;
				ELSIF rTemp_MovePos_M>rTemp_MovePos_G THEN
					i_plrTargetPos_All^:= i_plrTargetPos_All^-(rTemp_MovePos_G);
					i_plrTargetPos_M^:= i_plrTargetPos_M^-(rTemp_MovePos_M-rTemp_MovePos_G);
				ELSIF rTemp_MovePos_M<rTemp_MovePos_G THEN
					i_plrTargetPos_All^:= i_plrTargetPos_All^-(rTemp_MovePos_M);
					i_plrTargetPos_G^:= i_plrTargetPos_G^-(rTemp_MovePos_G-rTemp_MovePos_M);
				END_IF
			END_IF
		END_IF

		IF i_pstStTrapAxisParam_Gantray^.xFlag_MoveEn THEN
			IF i_pstStTrapAxisParam_Gantray^.lrPos_HandWheelChange<>0 THEN
				o_rVel:= ABS(i_pstStTrapAxisParam_Gantray^.lrPos_HandWheelChange*0.005*GC_LRMOTORPPR_TRAP*
					UINT_TO_REAL(i_uiNum)/
					i_rScrewPitch/
					UINT_TO_REAL(i_uiDen)/gc_TENSION_TSK_CYCLE_TIME);//*1.05;

				IF i_pstStTrapAxisParam_Gantray^.bySts_HandWheel=1 THEN
					i_plrTargetPos_All^:= i_plrTargetPos_All^-i_pstStTrapAxisParam_Gantray^.lrPos_HandWheelChange*0.005*GC_LRMOTORPPR_TRAP*
						UINT_TO_REAL(i_uiNum)/
						i_rScrewPitch/
						UINT_TO_REAL(i_uiDen);

				ELSIF i_pstStTrapAxisParam_Gantray^.bySts_HandWheel=2 THEN
					i_plrTargetPos_M^:= i_plrTargetPos_M^-i_pstStTrapAxisParam_Gantray^.lrPos_HandWheelChange*0.005*GC_LRMOTORPPR_TRAP*
						UINT_TO_REAL(i_uiNum)/
						i_rScrewPitch/
						UINT_TO_REAL(i_uiDen);

				ELSIF i_pstStTrapAxisParam_Gantray^.bySts_HandWheel=3 THEN
					i_plrTargetPos_G^:= i_plrTargetPos_G^-i_pstStTrapAxisParam_Gantray^.lrPos_HandWheelChange*0.005*GC_LRMOTORPPR_TRAP*
						UINT_TO_REAL(i_uiNum)/
						i_rScrewPitch/
						UINT_TO_REAL(i_uiDen);

				END_IF
			END_IF
		END_IF
(*
		IF i_pstStTrapAxisParam_Gantray^.xPressFlag_Stop  OR (i_pstStTrapAxisParam_Gantray^.xManuNeedStop AND i_pstStTrapAxisParam_Gantray^.xManuForPanel) THEN
			o_rVel:= 0;
			o_lrTargetPos_All:= i_pstStTrapAxisParam_Gantray^.lrPos_CurPos_Prf;
			o_lrTargetPos_M:= i_pstStTrapAxisParam_Gantray^.lrPos_CurPos_Prf_M;
			o_lrTargetPos_G:= i_pstStTrapAxisParam_Gantray^.lrPos_CurPos_Prf_G;
			IF i_pstStTrapAxisParam_Gantray^.xRev_Motor_M THEN
				i_plrTargetPos_All^:= -i_pstStTrapAxisParam_Gantray^.lrPos_CurPos_Prf;
				i_plrTargetPos_M^:= -i_pstStTrapAxisParam_Gantray^.lrPos_CurPos_Prf_M;
			ELSE
				i_plrTargetPos_All^:= i_pstStTrapAxisParam_Gantray^.lrPos_CurPos_Prf;
				i_plrTargetPos_M^:= i_pstStTrapAxisParam_Gantray^.lrPos_CurPos_Prf_M;
			END_IF
			IF i_pstStTrapAxisParam_Gantray^.xRev_Motor_G THEN
				i_plrTargetPos_G^:= -i_pstStTrapAxisParam_Gantray^.lrPos_CurPos_Prf_G;
			ELSE
				i_plrTargetPos_G^:= i_pstStTrapAxisParam_Gantray^.lrPos_CurPos_Prf_G;
			END_IF
		ELSE
			;
		END_IF
*)

		//2026.05.10.003923 | + | 增加限位保护,备份原来的位置
		//2026.05.10.003923 | + | 增加限位保护

		IF i_pstStTrapAxisParam_Gantray^.xPressFlag_Stop  OR (i_pstStTrapAxisParam_Gantray^.xManuNeedStop AND i_pstStTrapAxisParam_Gantray^.xManuForPanel) THEN
			rErr_TarPos_All := i_plrTargetPos_All^-rLast_TarPos_All;
			rErr_TarPos_M := i_plrTargetPos_M^ - rLast_TarPos_M;
			rErr_TarPos_G := i_plrTargetPos_G^ - rLast_TarPos_G;
			rErr_Pos := i_plrTargetPos_M^ - i_plrTargetPos_G^;

			IF i_pstStTrapAxisParam_Gantray^.lrParallelError_MM > i_rMaxErr THEN
				IF rErr_TarPos_M < 0 THEN
					o_rVel:= 0;
					i_plrTargetPos_All^:= rLast_TarPos_All;
					i_plrTargetPos_M^:= rLast_TarPos_M;
					i_plrTargetPos_G^:= rLast_TarPos_G;
				END_IF
				IF rErr_TarPos_G > 0 THEN
					o_rVel:= 0;
					i_plrTargetPos_All^:= rLast_TarPos_All;
					i_plrTargetPos_M^:= rLast_TarPos_M;
					i_plrTargetPos_G^:= rLast_TarPos_G;
				END_IF
			ELSIF i_pstStTrapAxisParam_Gantray^.lrParallelError_MM <-1*i_rMaxErr THEN
				IF rErr_TarPos_M > 0 THEN
					o_rVel:= 0;
					i_plrTargetPos_All^:= rLast_TarPos_All;
					i_plrTargetPos_M^:= rLast_TarPos_M;
					i_plrTargetPos_G^:= rLast_TarPos_G;
				END_IF
				IF rErr_TarPos_G < 0 THEN
					o_rVel:= 0;
					i_plrTargetPos_All^:= rLast_TarPos_All;
					i_plrTargetPos_M^:= rLast_TarPos_M;
					i_plrTargetPos_G^:= rLast_TarPos_G;
				END_IF

			END_IF
		ELSE
			rLast_TarPos_All := i_plrTargetPos_All^;
			rLast_TarPos_M := i_plrTargetPos_M^;
			rLast_TarPos_G := i_plrTargetPos_G^;
			rLast_ErrPos := rLast_TarPos_M - rLast_TarPos_G;
// 			IF ABS(rErr_Pos) > ABS(rLast_ErrPos) THEN
// 				o_rVel:= 0;
// 				o_lrTargetPos_All:= rLast_TarPos_All;
// 				o_lrTargetPos_M:= rLast_TarPos_M;
// 				o_lrTargetPos_G:= rLast_TarPos_G;
// 			ELSE
// 				;
// 			END_IF

		END_IF

		o_lrTargetPos_All:= i_plrTargetPos_All^;
		o_lrTargetPos_M:= i_plrTargetPos_M^;
		o_lrTargetPos_G:= i_plrTargetPos_G^;
		IF i_pstStTrapAxisParam_Gantray^.xRev_Motor_M THEN
			o_lrTargetPos_All:= -i_plrTargetPos_All^;
			o_lrTargetPos_M:= -i_plrTargetPos_M^;
		END_IF
		IF i_pstStTrapAxisParam_Gantray^.xRev_Motor_G THEN
			o_lrTargetPos_G:= -i_plrTargetPos_G^;
		END_IF

		//2026.05.10.003923 | + | 增加限位保护
// 		IF i_pstStTrapAxisParam_Gantray^.xPressFlag_Stop  OR (i_pstStTrapAxisParam_Gantray^.xManuNeedStop AND i_pstStTrapAxisParam_Gantray^.xManuForPanel) THEN
// 			rErr_TarPos_All := o_lrTargetPos_All-rLast_TarPos_All;
// 			rErr_TarPos_M := o_lrTargetPos_M - rLast_TarPos_M;
// 			rErr_TarPos_G := o_lrTargetPos_G - rLast_TarPos_G;
// 			rErr_Pos := o_lrTargetPos_M - o_lrTargetPos_G;
// 			IF ABS(rErr_Pos) > ABS(rLast_ErrPos) THEN
// 				o_rVel:= 0;
// 				o_lrTargetPos_All:= rLast_TarPos_All;
// 				o_lrTargetPos_M:= rLast_TarPos_M;
// 				o_lrTargetPos_G:= rLast_TarPos_G;
// 			ELSE
// 				;
// 			END_IF
// 		END_IF

		//处理标定模式下
		IF i_pstStTrapAxisParam_Gantray^.xSts_Calid_Pos THEN
			fbTRIG_Confirm_load_unload(CLK:=i_pstStTrapAxisParam_Gantray^.xConfirm_Load_Unload_Press);
			fbTRIG_Confirm_PressUp(CLK:=i_pstStTrapAxisParam_Gantray^.xConfirm_Up_Press);
			fbTRIG_Confirm_PressDn(CLK:=i_pstStTrapAxisParam_Gantray^.xConfirm_Dn_Press);
			i_pstStTrapAxisParam_Gantray^.xConfirm_Load_Unload_Press:= FALSE;
			i_pstStTrapAxisParam_Gantray^.xConfirm_Up_Press:= FALSE;
			i_pstStTrapAxisParam_Gantray^.xConfirm_Dn_Press:= FALSE;
			IF fbTRIG_Confirm_PressDn.Q THEN
				i_pstStTrapAxisParam_Gantray^.lrposConfirm_Dn_Press_M_Confirm:=
					i_pstStTrapAxisParam_Gantray^.lrPos_CurPos_Enc_M;
				i_pstStTrapAxisParam_Gantray^.lrposConfirm_Dn_Press_G_Confirm:=
					i_pstStTrapAxisParam_Gantray^.lrPos_CurPos_Enc_G;
				lrTemp:= i_rUp_Dn_Length*GC_LRMOTORPPR_TRAP*
						UINT_TO_REAL(i_uiNum)/
						i_rScrewPitch/
						UINT_TO_REAL(i_uiDen);
				g_lrtest:=lrTemp;
				IF 	i_pstStTrapAxisParam_Gantray^.xRev_Motor_M THEN
					i_pstStTrapAxisParam_Gantray^.lrposConfirm_Up_Press_M_Confirm:=
						i_pstStTrapAxisParam_Gantray^.lrposConfirm_Dn_Press_M_Confirm-lrTemp;
				ELSE
					i_pstStTrapAxisParam_Gantray^.lrposConfirm_Up_Press_M_Confirm:=
						i_pstStTrapAxisParam_Gantray^.lrposConfirm_Dn_Press_M_Confirm+lrTemp;
				END_IF
				IF 	i_pstStTrapAxisParam_Gantray^.xRev_Motor_G THEN
					i_pstStTrapAxisParam_Gantray^.lrposConfirm_Up_Press_G_Confirm:=
						i_pstStTrapAxisParam_Gantray^.lrposConfirm_Dn_Press_G_Confirm-lrTemp;
				ELSE
					i_pstStTrapAxisParam_Gantray^.lrposConfirm_Up_Press_G_Confirm:=
						i_pstStTrapAxisParam_Gantray^.lrposConfirm_Dn_Press_G_Confirm+lrTemp;
				END_IF
				//在这里记录一下标定时候的周长，秦华记录带长，只对于张带辊有效
				i_prGirth_Confirm^:= i_rGirth_Roller;
				i_pstStTrapAxisParam_Gantray^.xConfirmDnPosDne_Pressure_M := TRUE;//bai.zy | 2024.01.15.101452 | 标定完成标志
				i_pstStTrapAxisParam_Gantray^.xConfirmDnPosDne_Pressure_G := TRUE;//bai.zy | 2024.01.15.101452 | 标定完成标志
			END_IF
			IF fbTRIG_Confirm_load_unload.Q THEN
				i_pstStTrapAxisParam_Gantray^.lrposConfirm_Load_Unload_Press_M_Confirm:=
					i_pstStTrapAxisParam_Gantray^.lrPos_CurPos_Enc_M;
				i_pstStTrapAxisParam_Gantray^.lrposConfirm_Load_Unload_Press_G_Confirm:=
					i_pstStTrapAxisParam_Gantray^.lrPos_CurPos_Enc_G;
				i_pstStTrapAxisParam_Gantray^.xConfirmload_unloadPosDne_Pressure_M := TRUE;//bai.zy | 2024.01.15.101452 | 标定完成标志
				i_pstStTrapAxisParam_Gantray^.xConfirmload_unloadPosDne_Pressure_G := TRUE;//bai.zy | 2024.01.15.101452 | 标定完成标志
			END_IF
		ELSE//运行模式下可以矫正位置
			IF i_xFlag_Print AND
				(i_pstStTrapAxisParam_Gantray^.byCurPos_M=1 OR
				i_pstStTrapAxisParam_Gantray^.byCurPos_M=2 OR
				i_pstStTrapAxisParam_Gantray^.byCurPos_M=3) AND
				(i_pstStTrapAxisParam_Gantray^.byCurPos_G=1 OR
				i_pstStTrapAxisParam_Gantray^.byCurPos_G=2 OR
				i_pstStTrapAxisParam_Gantray^.byCurPos_G=3) (*AND
				i_pstStTrapAxisParam_Gantray^.xMove_To_Dn_Press_end*) THEN
				IF i_pstStTrapAxisParam_Gantray^.xConfirm_Adjust_PressDn OR //手轮按键矫正
						g_xConfirm_Adjust_PressDn THEN
					IF 	i_pstStTrapAxisParam_Gantray^.iStationId_M < 120 AND
						i_pstStTrapAxisParam_Gantray^.iStationId_G < 120 THEN

						lrTemp_Len_Load_Unload_Pos:= ABS(i_pstStTrapAxisParam_Gantray^.lrposConfirm_Dn_Press_M-
								i_pstStTrapAxisParam_Gantray^.lrposConfirm_Load_Unload_Press_M);

						i_pstStTrapAxisParam_Gantray^.lrposConfirm_Dn_Press_M_Confirm:=
							i_pstStTrapAxisParam_Gantray^.lrPos_CurPos_Enc_M;
						i_pstStTrapAxisParam_Gantray^.lrposConfirm_Dn_Press_G_Confirm:=
							i_pstStTrapAxisParam_Gantray^.lrPos_CurPos_Enc_G;

						lrTemp:= i_rUp_Dn_Length*GC_LRMOTORPPR_TRAP*
							UINT_TO_REAL(i_uiNum)/
							i_rScrewPitch/
							UINT_TO_REAL(i_uiDen);
						IF 	i_pstStTrapAxisParam_Gantray^.xRev_Motor_M THEN
							i_pstStTrapAxisParam_Gantray^.lrposConfirm_Up_Press_M_Confirm:=
								i_pstStTrapAxisParam_Gantray^.lrposConfirm_Dn_Press_M_Confirm-lrTemp;
							i_pstStTrapAxisParam_Gantray^.lrposConfirm_Load_Unload_Press_M_Confirm:=
								i_pstStTrapAxisParam_Gantray^.lrposConfirm_Dn_Press_M_Confirm-lrTemp_Len_Load_Unload_Pos;

						ELSE
							i_pstStTrapAxisParam_Gantray^.lrposConfirm_Up_Press_M_Confirm:=
								i_pstStTrapAxisParam_Gantray^.lrposConfirm_Dn_Press_M_Confirm+lrTemp;
							i_pstStTrapAxisParam_Gantray^.lrposConfirm_Load_Unload_Press_M_Confirm:=
								i_pstStTrapAxisParam_Gantray^.lrposConfirm_Dn_Press_M_Confirm+lrTemp_Len_Load_Unload_Pos;

						END_IF
						IF 	i_pstStTrapAxisParam_Gantray^.xRev_Motor_G THEN
							i_pstStTrapAxisParam_Gantray^.lrposConfirm_Up_Press_G_Confirm:=
								i_pstStTrapAxisParam_Gantray^.lrposConfirm_Dn_Press_G_Confirm-lrTemp;
							i_pstStTrapAxisParam_Gantray^.lrposConfirm_Load_Unload_Press_G_Confirm:=
								i_pstStTrapAxisParam_Gantray^.lrposConfirm_Dn_Press_G_Confirm-lrTemp_Len_Load_Unload_Pos;

						ELSE
							i_pstStTrapAxisParam_Gantray^.lrposConfirm_Up_Press_G_Confirm:=
								i_pstStTrapAxisParam_Gantray^.lrposConfirm_Dn_Press_G_Confirm+lrTemp;
							i_pstStTrapAxisParam_Gantray^.lrposConfirm_Load_Unload_Press_G_Confirm:=
								i_pstStTrapAxisParam_Gantray^.lrposConfirm_Dn_Press_G_Confirm+lrTemp_Len_Load_Unload_Pos;
						END_IF

						o_lrTemp_Len_Up_Pos := lrTemp;
						o_lrTemp_Len_Load_Unload_Pos := lrTemp_Len_Load_Unload_Pos;
						//在这里更新一下矫正时候的周长
						i_prGirth_Confirm^:= i_rGirth_Roller;
						i_pxFinishConfirm_Adjust_PressDn^ := TRUE;
					END_IF
				END_IF
			ELSE
				;
			END_IF
		END_IF
//2023.11.21.183755新增急停保护
		IF NOT i_pstStTrapAxisParam_Gantray^.xFlag_MoveEn OR (i_xFlag_Estop(* AND (NOT i_xMove_to_Up_Estop)*)) THEN//下私服需要重新处理一下输出2023.11.3.111425
			o_rVel:= 0;
			o_lrTargetPos_All:= i_pstStTrapAxisParam_Gantray^.lrPos_CurPos_Prf;
			o_lrTargetPos_M:= i_pstStTrapAxisParam_Gantray^.lrPos_CurPos_Prf_M;
			o_lrTargetPos_G:= i_pstStTrapAxisParam_Gantray^.lrPos_CurPos_Prf_G;
			IF i_pstStTrapAxisParam_Gantray^.xRev_Motor_M THEN
				i_plrTargetPos_All^:= -i_pstStTrapAxisParam_Gantray^.lrPos_CurPos_Prf;
				i_plrTargetPos_M^:= -i_pstStTrapAxisParam_Gantray^.lrPos_CurPos_Prf_M;
			ELSE
				i_plrTargetPos_All^:= i_pstStTrapAxisParam_Gantray^.lrPos_CurPos_Prf;
				i_plrTargetPos_M^:= i_pstStTrapAxisParam_Gantray^.lrPos_CurPos_Prf_M;
			END_IF
			IF i_pstStTrapAxisParam_Gantray^.xRev_Motor_G THEN
				i_plrTargetPos_G^:= -i_pstStTrapAxisParam_Gantray^.lrPos_CurPos_Prf_G;
			ELSE
				i_plrTargetPos_G^:= i_pstStTrapAxisParam_Gantray^.lrPos_CurPos_Prf_G;
			END_IF

			//2026.04.29.140841 | + | 急停或者下伺服状态把标志全清了
			i_pstStTrapAxisParam_Gantray^.xCanReFlashPos := FALSE;
			i_pstStTrapAxisParam_Gantray^.xRefleshPos := FALSE;
			i_pstStTrapAxisParam_Gantray^.xMove_To_PressDn := FALSE;
			i_pstStTrapAxisParam_Gantray^.xMove_To_PressUp := FALSE;
			i_pstStTrapAxisParam_Gantray^.xMove_To_Load_Unload := FALSE;

			//2026.05.08.130137 | + | 急停或者没有使能清标志
			i_pstStTrapAxisParam_Gantray^.xMove_To_Load_Unload_Press_ing:= FALSE;
			i_pstStTrapAxisParam_Gantray^.xMove_To_Up_Press_ing:= FALSE;
			i_pstStTrapAxisParam_Gantray^.xMove_To_Dn_Press_ing:= FALSE;
		END_IF

		//记录平行位置
		fbTRIG_Confirm_ParallelPos(CLK:=i_pstStTrapAxisParam_Gantray^.xConfirmParallelPos);
		IF fbTRIG_Confirm_ParallelPos.Q THEN
			i_pstStTrapAxisParam_Gantray^.lrEncPosParallel_M :=  i_pstStTrapAxisParam_Gantray^.lrPos_CurPos_Enc_M;
			i_pstStTrapAxisParam_Gantray^.lrEncPosParallel_G :=  i_pstStTrapAxisParam_Gantray^.lrPos_CurPos_Enc_G;
		END_IF

		//计算平行误差
		IF i_pstStTrapAxisParam_Gantray^.xRev_Motor_M AND i_pstStTrapAxisParam_Gantray^.lrEncPosParallel_M<>0 THEN
			lrEncParallelError_M := i_pstStTrapAxisParam_Gantray^.lrPos_CurPos_Enc_M - 1(*i_pstStTrapAxisParam_Gantray^.lrEncPosParallel_M*);

		ELSE
			lrEncParallelError_M := 1(*i_pstStTrapAxisParam_Gantray^.lrEncPosParallel_M*) - i_pstStTrapAxisParam_Gantray^.lrPos_CurPos_Enc_M;

		END_IF

		IF i_pstStTrapAxisParam_Gantray^.xRev_Motor_G AND i_pstStTrapAxisParam_Gantray^.lrEncPosParallel_G <> 0 THEN
			lrEncParallelError_G := i_pstStTrapAxisParam_Gantray^.lrPos_CurPos_Enc_G - 1(*i_pstStTrapAxisParam_Gantray^.lrEncPosParallel_G*);

		ELSE
			lrEncParallelError_G := 1(*i_pstStTrapAxisParam_Gantray^.lrEncPosParallel_G*) - i_pstStTrapAxisParam_Gantray^.lrPos_CurPos_Enc_G;

		END_IF

		IF i_rProportion <> 0 THEN
// 			i_pstStTrapAxisParam_Gantray^.lrParallelError_MM :=ABS((lrEncParallelError_M-lrEncParallelError_G)*
// 					i_rScrewPitch*UINT_TO_LREAL(i_uiDen)/GC_LRMOTORPPR_TRAP/UINT_TO_REAL(i_uiNum))/i_rProportion;
			i_pstStTrapAxisParam_Gantray^.lrParallelError_MM :=(lrEncParallelError_M-lrEncParallelError_G)*
				i_rScrewPitch*UINT_TO_LREAL(i_uiDen)/GC_LRMOTORPPR_TRAP/UINT_TO_REAL(i_uiNum)/i_rProportion;

		END_IF

		IF i_xFlag_Print AND
			(i_pstStTrapAxisParam_Gantray^.byCurPos_M=1 OR
			i_pstStTrapAxisParam_Gantray^.byCurPos_M=2 OR
			i_pstStTrapAxisParam_Gantray^.byCurPos_M=3) AND
			(i_pstStTrapAxisParam_Gantray^.byCurPos_G=1 OR
			i_pstStTrapAxisParam_Gantray^.byCurPos_G=2 OR
			i_pstStTrapAxisParam_Gantray^.byCurPos_G=3) AND
			i_pstStTrapAxisParam_Gantray^.xCanReFlashPos AND
			i_pstStTrapAxisParam_Gantray^.xRefleshPos THEN

			i_pstStTrapAxisParam_Gantray^.lrPrintPosOffsetDn_M:= i_pstStTrapAxisParam_Gantray^.lrCurPos_mm_M;
			i_pstStTrapAxisParam_Gantray^.lrPrintPosOffsetDn_G:= i_pstStTrapAxisParam_Gantray^.lrCurPos_mm_G;
			i_pstStTrapAxisParam_Gantray^.xCanReFlashPos := FALSE;
			i_pstStTrapAxisParam_Gantray^.xRefleshPos := FALSE;
		END_IF

		//记录最大限位
		fbTRIG_xCalidPressLimit_Max(CLK:=i_pstStTrapAxisParam_Gantray^.xCalidPressLimit_Max);
		IF fbTRIG_xCalidPressLimit_Max.Q THEN
			i_pstStTrapAxisParam_Gantray^.lrEncPosLimit_M_Max :=  i_pstStTrapAxisParam_Gantray^.lrPos_CurPos_Enc_M;
			i_pstStTrapAxisParam_Gantray^.lrEncPosLimit_G_Max :=  i_pstStTrapAxisParam_Gantray^.lrPos_CurPos_Enc_G;
		END_IF

		//在这里处理一下按钮功能；

	END_IF
END_IF

(* ---- KS_FB_McMultiFunCtl_GantryTrap.st ---- *)
(*@CES
Name=KS_FB_McMultiFunCtl_GantryTrap
Type=FunctionBlock
TypeGuid=6f9dac99-8de1-4efc-8465-68ac443b7d08
Guid=b1cd30ae-efbb-4f40-9386-b86c83b34233
HasDeclaration=True
HasImplementation=True
*)
{DECLARATION}
FUNCTION_BLOCK KS_FB_McMultiFunCtl_GantryTrap(*大指令控制*)
(*
1.检查伺服状态
2.大指令写控制
*)
VAR_INPUT
	i_xEn: BOOL;
	i_iGrpId: INT;
	i_iGrpGantryTrapGroup_Num: INT;
	i_iGrpGantryTrapMotion_Num: INT;
	i_aiGrpGantryTrapMotion_StdList: ARRAY [1..MAX_STATION_NUM] OF INT;
	i_pstStSysParam: POINTER TO StSysParam;
	i_pastStAxisIdListInf :POINTER TO ARRAY [1..128] OF StAxisIdListInf;
	i_pastStSetPrm					:POINTER TO ARRAY [1..MAX_STATION_NUM] OF TSetMultiMcFunctionPrm;
	i_pastStGetMotionSts: POINTER TO ARRAY [1..MAX_STATION_NUM] OF StGetMotionSts;
	i_pastStMotorParam_GantryTrap: POINTER TO ARRAY [1..MAX_STATION_NUM] OF StMotorParam_GantryTrap;
	i_pstStHYLogFifo			: POINTER TO StHYLogFifo;(* 2025.8.23.170701/han.dp/增加的日志队列 *)
END_VAR
VAR_OUTPUT
END_VAR
VAR_IN_OUT
END_VAR
VAR
	iN : INT;
	iRtn: INT;
	alrVarValue : ARRAY [1..80] OF LREAL;
	dwRtn : DWORD;
	astStSetPrm_Pre				: ARRAY [1..MAX_STATION_NUM] OF TSetMultiMcFunctionPrm;

	fbKS_FB_CheckServeOnDone_GantryTrap : KS_FB_CheckServeOnDone_GantryTrap;
	pstStGrpParam_Save : POINTER TO StGrpParam_Save;
	pstStGrpParam_UnSave : POINTER TO StGrpParam_UnSave;

	iRtn_McMulFun : INT ;
	iRtn_McMulFun_Pre : INT ;

	sTMultiMcFunctionReadPrm : TMultiMcFunctionReadPrm;

	(*2025-12-10 by sjw 非阻塞大指令*)
	FB_Set_StartMcMUltiFunction: GTMC_StartMcMultiFunction;
	bDoneSet: BOOL := TRUE;
	bBusySet: BOOL;
	bErrorSet: BOOL;
	iErrorIdSet: INT;
END_VAR

{IMPLEMENTATION}
(*1.伺服检查-确保所有需要转的轴都上伺服了才能进行下一步*)
pstStGrpParam_Save := ADR(i_pstStSysParam^.astStGrpParam_Save[i_iGrpId]);
pstStGrpParam_UnSave := ADR(i_pstStSysParam^.astStGrpParam_UnSave[i_iGrpId]);

fbKS_FB_CheckServeOnDone_GantryTrap(
	i_xEn:= ((pstStGrpParam_Save^.wCtl_Pressure_Up_Dn.5) AND (NOT fbKS_FB_CheckServeOnDone_GantryTrap.o_xDone)),
	i_iGrpGantryTrapGroup_Num := i_iGrpGantryTrapGroup_Num,
	i_iGrpGantryTrapMotion_Num:= i_iGrpGantryTrapMotion_Num,
	i_aiGrpGantryTrapMotion_StdList:= i_aiGrpGantryTrapMotion_StdList,
	i_pstStSysParam:= i_pstStSysParam,
	i_pastStAxisIdListInf:= i_pastStAxisIdListInf,
	i_pastStGetMotionSts:= i_pastStGetMotionSts,
	i_pastStMotorParam_GantryTrap:= i_pastStMotorParam_GantryTrap,
	i_xFlag_StopOrEStop := pstStGrpParam_UnSave^.xFlag_Stop OR pstStGrpParam_UnSave^.xFlag_Estop,
	o_xEn=> ,
	o_xDone=> ,
	o_iErrNo=> ,
	o_iErrAxisId=> ,
	o_iErrTypeId=> ,
	o_iErrUnitId=> ,
	o_iErrCoreId=> );

(*2.大指令写*)
sTMultiMcFunctionReadPrm.readCommandVarTableIndex := 1;
sTMultiMcFunctionReadPrm.readCount := 0;
sTMultiMcFunctionReadPrm.pVarValue := ADR(alrVarValue);
dwRtn:= SysMemCmp(i_pastStSetPrm,ADR(astStSetPrm_Pre),SIZEOF(astStSetPrm_Pre));
IF dwRtn<>0 THEN
	//修改非阻塞方式 2025-12-10 by sjw
	iRtn_McMulFun:=GTN_StartMcMultiFunction(2,INT_TO_UINT(i_iGrpGantryTrapGroup_Num),1,i_pastStSetPrm,ADR(sTMultiMcFunctionReadPrm));
	IF iRtn_McMulFun <> 0 AND iRtn_McMulFun_Pre <> iRtn_McMulFun THEN
		KS_HY_AddMsgToLog(g_pstStHYLogFifo, LOG_LEVEL_ALARM, 'GTN_StartMcMultiFunction GantryTrap Err!', INT_TO_STRING(iRtn_McMulFun));
	END_IF
	iRtn_McMulFun_Pre := iRtn_McMulFun;
	(*
	IF bDoneSet  = TRUE AND bBusySet = FALSE THEN
		FB_Set_StartMcMUltiFunction(
		Execute:= TRUE,
		Block:= TRUE,
		core:= 2,
		axisCount:= INT_TO_UINT(i_iGrpGantryTrapGroup_Num),
		writeEnable:= 1,
		pSetPrm:= i_pastStSetPrm,
		pGetPrm:= ADR(sTMultiMcFunctionReadPrm),
		Done=> bDoneSet,
		Busy=> bBusySet,
		Error=> bErrorSet,
		ErrorID=> iErrorIdSet);
	END_IF
	*)
END_IF
SysMemCpy(ADR(astStSetPrm_Pre),i_pastStSetPrm,SIZEOF(i_pastStSetPrm^));
